(* IEC 61131-3 sources: beedance/reference (part 10) *)

// Commented out for beedance: it uses CHR_TO_STRING, which is commented out.
// FUNCTION_BLOCK TN_INPUT_EDIT_LINE
// VAR
// 	in_count : INT;
// 	in_Count_End : INT;
// 	in_CursorOffset : INT;
// 	by_Attr : BYTE;
// 	st_String : STRING;
// 	bo_Pos_Found : BOOL;
// 	st_CHAR : STRING(1);
// 	in_old_charpos : INT;
// END_VAR
// VAR
// 	FB_TN_SC_WRITE : TN_SC_WRITE;
// END_VAR
// VAR_IN_OUT
// 	Xus_TN_SCREEN : us_TN_SCREEN;
// 	Xus_TN_INPUT_CONTROL_DATA : us_TN_INPUT_CONTROL_DATA;
// END_VAR
//
// (* Cursorsteuerung rücksetzen *)
// in_CursorOffset := INT#0;
//
// IF Xus_TN_INPUT_CONTROL_DATA.bo_Focus = TRUE THEN
//
// 	(* Texteingabe erkannt ? *)
// 	IF Xus_TN_INPUT_CONTROL_DATA.by_Input_ASCII_Code > BYTE#0 THEN
//
// 		IF (Xus_TN_INPUT_CONTROL_DATA.bo_Input_Only_Num = TRUE AND Xus_TN_INPUT_CONTROL_DATA.bo_Input_ASCII_IsNum = TRUE)
// 			OR (Xus_TN_INPUT_CONTROL_DATA.bo_Input_Only_Num = FALSE) THEN
//
// 			(* ASCII Wert in einen String wandeln *)
// 			st_CHAR := CHR_TO_STRING(C:=Xus_TN_INPUT_CONTROL_DATA.by_Input_ASCII_Code);
//
// 			(* Eingabe übernehmen *)
// 			Xus_TN_INPUT_CONTROL_DATA.st_Input_Data := REPLACE(Xus_TN_INPUT_CONTROL_DATA.st_Input_Data,
// 			st_CHAR,INT#1,Xus_TN_INPUT_CONTROL_DATA.in_Cursor_Pos);
//
// 			in_CursorOffset := INT#1;
// 			Xus_TN_INPUT_CONTROL_DATA.bo_Update_Input := TRUE;
// 		END_IF;
// 	END_IF;
//
// 	CASE BYTE_TO_INT(Xus_TN_INPUT_CONTROL_DATA.by_Input_Exten_Code) OF
//
// 	67: (* Cursor rechts gedrückt *)
// 		in_CursorOffset := INT#1;
//
// 	68: (* Cursor links gedrückt *)
// 		in_CursorOffset := -1;
//
// 	08: (* Backspace gedrückt *)
// 		Xus_TN_INPUT_CONTROL_DATA.st_Input_Data := REPLACE(Xus_TN_INPUT_CONTROL_DATA.st_Input_Data, ' ', 1,Xus_TN_INPUT_CONTROL_DATA.in_Cursor_Pos);
// 		Xus_TN_INPUT_CONTROL_DATA.bo_Update_Input := TRUE;
// 		in_CursorOffset := -1;
//
// 	13: (* Enter-Taste gedrückt *)
// 		IF LEN(Xus_TN_INPUT_CONTROL_DATA.st_Input_Mask) > INT#00 THEN
// 			(* Eingabestring übernehmen *)
// 			Xus_TN_INPUT_CONTROL_DATA.st_Input_String := Xus_TN_INPUT_CONTROL_DATA.st_Input_Data;
//
// 			(* Eingabestring -> links und rechts Leerzeichen entfernen *)
// 			Xus_TN_INPUT_CONTROL_DATA.st_Input_String := TRIME(str:=Xus_TN_INPUT_CONTROL_DATA.st_Input_String);
// 			Xus_TN_INPUT_CONTROL_DATA.bo_Input_Entered := TRUE;
//
// 			(* neue Eingabe vorbereiten *)
// 			Xus_TN_INPUT_CONTROL_DATA.st_Input_Data := Xus_TN_INPUT_CONTROL_DATA.st_Input_Mask;
//
// 			Xus_TN_INPUT_CONTROL_DATA.in_Cursor_Pos := INT#1;
// 			Xus_TN_INPUT_CONTROL_DATA.bo_Update_Input := TRUE;
//
// 			(* suche erstes Position in Eingabemaske *)
// 			st_CHAR := MID(Xus_TN_INPUT_CONTROL_DATA.st_Input_Mask,1,Xus_TN_INPUT_CONTROL_DATA.in_Cursor_Pos);
// 			IF st_CHAR <> ' ' THEN
// 				(* nächsten Eingabeposition suchen *)
// 				in_CursorOffset := INT#1;
// 			END_IF;
// 		END_IF;
// 	END_CASE;
// END_IF;
//
// (* Cursor richtung rechts bewegen                                   *)
// IF (in_CursorOffset > INT#0) OR (Xus_TN_INPUT_CONTROL_DATA.in_Cursor_Pos = INT#0) THEN
// 	bo_Pos_Found := FALSE;
//
// 	in_Count := Xus_TN_INPUT_CONTROL_DATA.in_Cursor_Pos + INT#1;
// 	in_Count_End := LEN(Xus_TN_INPUT_CONTROL_DATA.st_Input_Mask);
//
// 	WHILE (in_count <= in_Count_End) AND (bo_Pos_Found = FALSE) DO
//
// 		st_CHAR := MID(Xus_TN_INPUT_CONTROL_DATA.st_Input_Mask,1,in_count);
// 		IF st_CHAR = ' ' THEN
// 			Xus_TN_INPUT_CONTROL_DATA.in_Cursor_Pos := in_count;
// 			Xus_TN_INPUT_CONTROL_DATA.bo_Update_Input := TRUE;
// 			bo_Pos_Found := TRUE;
// 		END_IF;
//
// 		in_count := in_count + INT#1;
//
// 	END_WHILE;
// END_IF;
//
// (* Cursor richtung links bewegen *)
// IF in_CursorOffset < INT#0 THEN
// 	bo_Pos_Found := FALSE;
//
// 	in_Count     := Xus_TN_INPUT_CONTROL_DATA.in_Cursor_Pos - INT#01;
// 	in_Count_End := INT#1;
//
// 	WHILE (in_count >= in_Count_End) AND (bo_Pos_Found = FALSE) DO
//
// 		st_CHAR := MID(Xus_TN_INPUT_CONTROL_DATA.st_Input_Mask,1,in_count);
// 		IF st_CHAR = ' ' THEN
// 			Xus_TN_INPUT_CONTROL_DATA.in_Cursor_Pos := in_count;
// 			Xus_TN_INPUT_CONTROL_DATA.bo_Update_Input := TRUE;
// 			bo_Pos_Found := TRUE;
// 		END_IF;
//
// 		in_count := in_count - INT#1;
// 	END_WHILE;
// END_IF;
//
// (* maximale Cursorposition ? *)
// IF Xus_TN_INPUT_CONTROL_DATA.in_Cursor_Pos > LEN(Xus_TN_INPUT_CONTROL_DATA.st_Input_Data) THEN
// 	Xus_TN_INPUT_CONTROL_DATA.in_Cursor_Pos := LEN(Xus_TN_INPUT_CONTROL_DATA.st_Input_Data);
// 	Xus_TN_INPUT_CONTROL_DATA.bo_Update_Input := TRUE;
// END_IF;
//
// (* minimale Cursorposition ? *)
// IF Xus_TN_INPUT_CONTROL_DATA.in_Cursor_Pos < INT#1 THEN
// 	Xus_TN_INPUT_CONTROL_DATA.in_Cursor_Pos := INT#1;
// 	Xus_TN_INPUT_CONTROL_DATA.bo_Update_Input := TRUE;
// END_IF;
//
// (* Aktualisierung der Anzeige *)
// IF (Xus_TN_INPUT_CONTROL_DATA.bo_Update_Input = TRUE) OR (Xus_TN_INPUT_CONTROL_DATA.bo_Update_All = TRUE) THEN
//
// 	(* Title-Text ausgeben *)
// 	IF (Xus_TN_INPUT_CONTROL_DATA.bo_Update_All = TRUE) THEN
//
// 		IF (Xus_TN_INPUT_CONTROL_DATA.in_Title_X_Offset = INT#00) AND (Xus_TN_INPUT_CONTROL_DATA.in_Title_Y_Offset = INT#00) THEN
// 			(* wenn Offset X,Y =0 dann Titlestring links vom Element positionieren *)
// 			FB_TN_SC_WRITE.Iin_Y := Xus_TN_INPUT_CONTROL_DATA.in_Y;
// 			FB_TN_SC_WRITE.Iin_X := Xus_TN_INPUT_CONTROL_DATA.in_X - LEN(Xus_TN_INPUT_CONTROL_DATA.st_Title_String);
// 		ELSE
// 			(* Title-Text durch Row, Color-Offset ausgeben *)
// 			FB_TN_SC_WRITE.Iin_Y := Xus_TN_INPUT_CONTROL_DATA.in_Y + Xus_TN_INPUT_CONTROL_DATA.in_Title_Y_Offset;
// 			FB_TN_SC_WRITE.Iin_X := Xus_TN_INPUT_CONTROL_DATA.in_X + Xus_TN_INPUT_CONTROL_DATA.in_Title_X_Offset;
// 		END_IF;
//
// 		(* Title-Text durch Row, Color-Offset ausgeben *)
// 		FB_TN_SC_WRITE(	Iby_ATTR := Xus_TN_INPUT_CONTROL_DATA.by_Title_Attr,
// 						Ist_STRING := Xus_TN_INPUT_CONTROL_DATA.st_Title_String,
// 						Xus_TN_SCREEN := Xus_TN_SCREEN);
// 	END_IF;
//
// 	(* Eingabetext ausgeben *)
// 	IF (Xus_TN_INPUT_CONTROL_DATA.bo_Input_Hidden = TRUE) THEN
//
// 		st_String := '';
//
// 		IF LEN(Xus_TN_INPUT_CONTROL_DATA.st_Input_Data) = LEN(Xus_TN_INPUT_CONTROL_DATA.st_Input_Mask) THEN
// 			(* Eingabemodus: HIDDEN *)
// 			FOR in_count := 1 TO LEN(Xus_TN_INPUT_CONTROL_DATA.st_Input_Data) DO
//
// 				(* Zeichen aus Eingabemaske lesen *)
// 				st_CHAR := MID(Xus_TN_INPUT_CONTROL_DATA.st_Input_Mask,1,in_count);
//
// 				(* Eingabe oder Maskenzeichen ausgeben *)
// 				IF st_CHAR = ' ' THEN
//
// 					(* Zeichen aus Eingabedata lesen *)
// 					st_CHAR := MID(Xus_TN_INPUT_CONTROL_DATA.st_Input_Data,1,in_count);
//
// 					IF st_CHAR = ' ' THEN
// 						(* Leerzeichen ausgeben *)
// 						st_String := CONCAT(st_String, ' ');
//
// 					ELSE
// 						(* verdecktes Zeichen ausgeben *)
// 						st_String := CONCAT(st_String, '*');
//
// 					END_IF;
//
// 				ELSE
// 					(* Zeichen aus Eingabemaske übernehmen *)
// 					st_CHAR := MID(Xus_TN_INPUT_CONTROL_DATA.st_Input_Data,1,in_count);
// 					st_String := CONCAT(st_String,st_CHAR);
//
// 				END_IF;
// 			END_FOR;
// 		END_IF;
// 	ELSE
//
// 		(* Eingabemodus: NORMAL *)
// 		st_String := Xus_TN_INPUT_CONTROL_DATA.st_Input_Data;
//
// 	END_IF;
//
// 	(* String ausgeben *)
//
// 	IF Xus_TN_INPUT_CONTROL_DATA.bo_Focus = TRUE THEN
// 		by_Attr := Xus_TN_INPUT_CONTROL_DATA.by_Attr_mF;
// 	ELSE
// 		by_Attr := Xus_TN_INPUT_CONTROL_DATA.by_Attr_oF;
// 	END_IF;
//
// 	FB_TN_SC_WRITE(	Iin_Y := Xus_TN_INPUT_CONTROL_DATA.in_Y,
// 					Iin_X := Xus_TN_INPUT_CONTROL_DATA.in_X,
// 					Iby_ATTR := by_Attr,
// 					Ist_STRING := st_String,
// 					Xus_TN_SCREEN := Xus_TN_SCREEN);
//
// 	(* Cursor auf aktuelle Position setzen *)
// 	Xus_TN_INPUT_CONTROL_DATA.in_Cursor_Y := Xus_TN_INPUT_CONTROL_DATA.in_Y;
// 	Xus_TN_INPUT_CONTROL_DATA.in_Cursor_X := Xus_TN_INPUT_CONTROL_DATA.in_X + Xus_TN_INPUT_CONTROL_DATA.in_Cursor_Pos - INT#1;
//
// 	in_old_charpos := INT#0;
//
// 	(* Update-Flag's rücksetzen *)
// 	Xus_TN_INPUT_CONTROL_DATA.bo_Update_All := FALSE;
// 	Xus_TN_INPUT_CONTROL_DATA.bo_Update_Input := FALSE;
// END_IF;
// END_FUNCTION_BLOCK

// Commented out for beedance: it uses ELEMENT_GET, which is commented out.
// FUNCTION_BLOCK TN_INPUT_MENU_BAR
// VAR
// 	FB_TN_INPUT_MENU_POPUP : TN_INPUT_MENU_POPUP;
// 	us_TN_MENU_POPUP : us_TN_MENU_POPUP;
// 	FB_TN_SC_WRITE_C : TN_SC_WRITE_C;
// END_VAR
// VAR
// 	in_ROW : INT;
// 	in_COL : INT;
// 	in_TITLE_Length : INT;
// 	st_MENU_BAR : STRING(STRING_LENGTH);
// 	st_MENU_TITLE : STRING;
// 	in_Count : INT;
// 	in_Index : INT;
// 	by_New_KeyCode : BYTE;
// 	in_Scroll_Offset : INT;
// 	by_ATTR : BYTE;
// 	bo_Reset_Position :	BOOL;
// END_VAR
// VAR_IN_OUT
// 	Xus_TN_MENU : us_TN_MENU;
// 	Xus_TN_SCREEN : us_TN_SCREEN;
// END_VAR
//
// (* sicherstellen das rechteck immer innerhalb screen positioniert wird *)
//
// IF (Xus_TN_MENU.in_State = INT#00) AND (Xus_TN_MENU.bo_Create = TRUE) THEN
// 	Xus_TN_MENU.in_State := INT#01;
// 	Xus_TN_MENU.bo_Create := FALSE;
// 	Xus_TN_MENU.in_Menu_Selected := INT#00;
// 	Xus_TN_MENU.bo_Update := TRUE;
// 	bo_Reset_Position := TRUE;
//
// 	(* Menu-Bar - Hauptmenue *)
// 	st_MENU_BAR := ELEMENT_GET(SEP:=BYTE#37,POS:=0,ELEMENT:=Xus_TN_MENU.st_MENU_TEXT);
//
// 	(* Menu-Bar - Anzahl der Elemente bestimmen *)
// 	Xus_TN_MENU.in_Menu_E_Count := ELEMENT_COUNT(SEP:=BYTE#35,ELEMENT:=st_MENU_BAR);
//
// END_IF;
//
// (* Keycode ablegen *)
// by_New_KeyCode := Xus_TN_SCREEN.by_Input_Exten_Code;
//
// (* Popup-Menu Tastensteuerung (nur Cursor oben + unten zulassen *)
// IF (by_New_KeyCode = BYTE#65) OR (by_New_KeyCode = BYTE#66) THEN
// 	us_TN_MENU_POPUP.by_Input_Exten_Code := by_New_KeyCode;
// ELSE
// 	us_TN_MENU_POPUP.by_Input_Exten_Code := BYTE#00;
// END_IF;
//
// (* Escape *)
// IF (by_New_KeyCode = BYTE#27) THEN
// 	(* Menu war inaktiv -> Escape -> Menu aktivieren *)
// 	IF (Xus_TN_MENU.in_State = INT#01) AND (Xus_TN_SCREEN.bo_Modal_Dialog = FALSE) THEN
// 		Xus_TN_MENU.in_State := INT#02;
// 		Xus_TN_MENU.bo_Update := TRUE;
// 		Xus_TN_MENU.in_Menu_Selected := INT#00;
//
// 		Xus_TN_SCREEN.bo_Menue_Bar_Dialog := TRUE;
//
// 		(* Menu war aktiv -> Escape -> Menu deaktivieren *)
// 	ELSIF (Xus_TN_MENU.in_State = INT#02) THEN
// 		us_TN_MENU_POPUP.bo_Destroy := TRUE;
// 		Xus_TN_MENU.bo_Update := TRUE;
// 		Xus_TN_MENU.in_State := INT#01;
// 		bo_Reset_Position := TRUE;
//
// 		Xus_TN_SCREEN.bo_Menue_Bar_Dialog := FALSE;
// 	END_IF;
// END_IF;
//
// (* Menu aktiv *)
// IF (Xus_TN_MENU.in_State = INT#02) THEN
//
// 	(* Return *)
// 	IF (by_New_KeyCode = BYTE#13)  THEN
// 		us_TN_MENU_POPUP.bo_Destroy := TRUE;
// 		Xus_TN_MENU.bo_Update := TRUE;
// 		Xus_TN_MENU.in_State := INT#01;
// 		bo_Reset_Position := TRUE;
// 		Xus_TN_MENU.in_Menu_Selected := (Xus_TN_MENU.in_Cur_Menu_Item * INT#10) + Xus_TN_MENU.in_Cur_Sub_Item;
// 		Xus_TN_SCREEN.by_Input_Exten_Code := BYTE#00;
//
// 		Xus_TN_SCREEN.bo_Menue_Bar_Dialog := FALSE;
//
// 		(* Destroy-Befehl -> Popup-Menu beenden *)
// 	ELSIF (Xus_TN_MENU.bo_Destroy = TRUE) THEN
// 		us_TN_MENU_POPUP.bo_Destroy := TRUE;
// 		Xus_TN_MENU.bo_Update := TRUE;
// 		Xus_TN_MENU.in_State := INT#01;
// 		bo_Reset_Position := TRUE;
// 		Xus_TN_MENU.in_Menu_Selected := INT#00;
// 		Xus_TN_SCREEN.by_Input_Exten_Code := BYTE#00;
//
// 		Xus_TN_SCREEN.bo_Menue_Bar_Dialog := FALSE;
//
// 	END_IF;
//
// 	IF (by_New_KeyCode = BYTE#67) THEN (* Cursor rechts *)
// 		in_Scroll_Offset := INT#1;
// 		Xus_TN_MENU.bo_Update := TRUE;
// 		Xus_TN_SCREEN.by_Input_Exten_Code := BYTE#00;
//
// 	ELSIF (by_New_KeyCode = BYTE#68) THEN (* Cursor links *)
// 		in_Scroll_Offset := -1;
// 		Xus_TN_MENU.bo_Update := TRUE;
// 		Xus_TN_SCREEN.by_Input_Exten_Code := BYTE#00;
// 	END_IF;
// END_IF;
//
// IF bo_Reset_Position = TRUE THEN
// 	bo_Reset_Position := FALSE;
// 	Xus_TN_MENU.in_X_SM_old := -1;
// 	Xus_TN_MENU.in_Y_SM_old := -1;
// 	Xus_TN_MENU.in_X_SM_new := -1;
// 	Xus_TN_MENU.in_Y_SM_new := -1;
// END_IF;
//
// (* POPUP-Menu updaten *)
// IF (Xus_TN_MENU.in_State > INT#00) AND (Xus_TN_MENU.bo_Update = TRUE) THEN
//
// 	Xus_TN_MENU.bo_Update := FALSE;
//
// 	in_ROW := Xus_TN_MENU.in_Y;
// 	in_COL := Xus_TN_MENU.in_X;
//
// 	(* Scrolloffset *)
// 	IF in_Scroll_Offset <> INT#00 THEN
// 		Xus_TN_MENU.in_Cur_Menu_Item := INC2(Xus_TN_MENU.in_Cur_Menu_Item,in_Scroll_Offset,1,Xus_TN_MENU.in_Menu_E_Count);
// 		in_Scroll_Offset := INT#00;
// 	ELSE
// 		(* Item = 0 und kein Scrolloffset *)
// 		IF (Xus_TN_MENU.in_Cur_Menu_Item = INT#00) THEN
// 			Xus_TN_MENU.in_Cur_Menu_Item := INT#01;
// 		END_IF;
// 	END_IF;
//
// 	(* alle Menutext zeichnen *)
// 	FOR in_Count := INT#01 TO Xus_TN_MENU.in_Menu_E_Count DO;
//
// 		(* Zeichenfarbe bestimmen *)
// 		IF (in_Count = Xus_TN_MENU.in_Cur_Menu_Item) AND (Xus_TN_MENU.in_State > INT#01 ) THEN
// 			by_ATTR := Xus_TN_MENU.by_Attr_mF;
//
// 			Xus_TN_MENU.in_Y_SM_new := in_ROW + INT#01;
// 			Xus_TN_MENU.in_X_SM_new := in_COL;
//
// 		ELSE
// 			by_ATTR := Xus_TN_MENU.by_Attr_oF;
// 		END_IF;
//
// 		st_MENU_TITLE := ELEMENT_GET(SEP:=BYTE#35,POS:=in_Count - 1,ELEMENT:=st_MENU_BAR);
//
// 		in_TITLE_Length := LEN(st_MENU_TITLE) + INT#02;
//
// 		FB_TN_SC_WRITE_C(	Iin_Y := in_ROW,
// 							Iin_X := in_COL,
// 							Iby_ATTR := by_ATTR,
// 							Iin_LENGTH := in_TITLE_Length,
// 							Iin_OPTION := INT#02,
// 							Ist_STRING := st_MENU_TITLE,
// 							Xus_TN_SCREEN := Xus_TN_SCREEN);
//
// 		in_COL := in_COL + in_TITLE_Length;
//
// 	END_FOR;
// END_IF;
//
// IF Xus_TN_MENU.in_X_SM_new <> Xus_TN_MENU.in_X_SM_old THEN
//
// 	(* SubMenu ist aktiv -> beenden                                     *)
// 	IF us_TN_MENU_POPUP.bo_Activ = TRUE THEN
// 		us_TN_MENU_POPUP.bo_Destroy := TRUE;
//
// 		(* Sub-Menu bearbeiten *)
// 		FB_TN_INPUT_MENU_POPUP(	Xus_TN_MENU_POPUP := us_TN_MENU_POPUP,
// 								Xus_TN_SCREEN := Xus_TN_SCREEN);
// 	END_IF;
//
// 	IF us_TN_MENU_POPUP.bo_Activ = FALSE THEN
// 		(* Popup-Menu zu aktuellen Menu parametrieren und ausführen         *)
// 		in_Index := Xus_TN_MENU.in_Cur_Menu_Item;
//
// 		us_TN_MENU_POPUP.in_Y := Xus_TN_MENU.in_Y_SM_new;
// 		us_TN_MENU_POPUP.in_X := Xus_TN_MENU.in_X_SM_new;
// 		us_TN_MENU_POPUP.by_Attr_mF := Xus_TN_MENU.by_Attr_mF;
// 		us_TN_MENU_POPUP.by_Attr_oF := Xus_TN_MENU.by_Attr_oF;
// 		us_TN_MENU_POPUP.st_Menu_Text := ELEMENT_GET(SEP:=BYTE#37,POS:=in_Index,ELEMENT:=Xus_TN_MENU.st_MENU_TEXT);
// 		us_TN_MENU_POPUP.bo_Create := TRUE;
//
// 		Xus_TN_MENU.in_X_SM_old := Xus_TN_MENU.in_X_SM_new;
// 		Xus_TN_MENU.in_Y_SM_old := Xus_TN_MENU.in_Y_SM_new;
//
// 	END_IF;
// END_IF;
//
// (* Popup-Menu zyklisch aufrufen *)
// FB_TN_INPUT_MENU_POPUP(	Xus_TN_MENU_POPUP := us_TN_MENU_POPUP,
// 						Xus_TN_SCREEN := Xus_TN_SCREEN);
//
// (* aktuelles Item vom Popup-Menu kopieren *)
// Xus_TN_MENU.in_Cur_Sub_Item := us_TN_MENU_POPUP.in_Cur_Item;
//
// (* Destroy-Befehl *)
// IF (Xus_TN_MENU.in_State = INT#01) THEN
// 	IF (Xus_TN_MENU.bo_Destroy = TRUE) THEN
// 		Xus_TN_MENU.in_State := INT#00;
// 		Xus_TN_MENU.bo_Destroy := FALSE;
// 		Xus_TN_MENU.in_Cur_Menu_Item := INT#00;
// 		Xus_TN_MENU.in_Cur_Sub_Item := INT#00;
// 	END_IF;
// END_IF;
// END_FUNCTION_BLOCK

// Commented out for beedance: it uses ELEMENT_COUNT, which is commented out.
// FUNCTION_BLOCK TN_INPUT_MENU_POPUP
// VAR
// 	FB_TN_SC_AREA_SAVE : TN_SC_AREA_SAVE;
// 	FB_TN_SC_AREA_RESTORE : TN_SC_AREA_RESTORE;
// 	FB_TN_SC_LINE : TN_SC_LINE;
// 	FB_TN_SC_ADD_SHADOW : TN_SC_ADD_SHADOW;
// 	FB_TN_SC_BOX : TN_SC_BOX;
// 	FB_TN_SC_WRITE_C : TN_SC_WRITE_C;
// END_VAR
// VAR
// 	in_ROW : INT;
// 	in_ROWS : INT;
// 	in_COL : INT;
// 	in_COLS : INT;
// 	in_index : INT;
// 	in_Count : INT;
// 	in_Scroll_Offset : INT;
// 	by_ATTR : BYTE;
// END_VAR
// VAR_IN_OUT
// 	Xus_TN_MENU_POPUP : us_TN_MENU_POPUP;
// 	Xus_TN_SCREEN : us_TN_SCREEN;
// END_VAR
//
// (* sicherstellen das rechteck immer innerhalb screen positioniert wird *)
//
// IF (Xus_TN_MENU_POPUP.bo_Activ = FALSE) AND (Xus_TN_MENU_POPUP.bo_Create = TRUE) THEN
// 	Xus_TN_MENU_POPUP.bo_Activ := TRUE;
// 	Xus_TN_MENU_POPUP.bo_Create := FALSE;
// 	Xus_TN_MENU_POPUP.bo_Destroy := FALSE;
// 	Xus_TN_MENU_POPUP.bo_Update := TRUE;
//
//   (* Sub-Menu-Texte *)
//
// 	Xus_TN_MENU_POPUP.in_Menu_E_Count := ELEMENT_COUNT(SEP:=BYTE#35,ELEMENT:=Xus_TN_MENU_POPUP.st_Menu_Text);
//
// 	(* Anzahl Zeilen (Sub-Menu-Texte) bestimmen *)
// 	Xus_TN_MENU_POPUP.in_Rows := Xus_TN_MENU_POPUP.in_Menu_E_Count;
//
// 	(* längsten Sub-Menu-Text suchen *)
// 	Xus_TN_MENU_POPUP.in_Cols := INT#00;
//
// 	FOR in_Count := INT#01 TO Xus_TN_MENU_POPUP.in_Rows DO;
// 		Xus_TN_MENU_POPUP.in_Cols:=MAX(LEN(ELEMENT_GET(SEP:=BYTE#35,POS:=in_Count - 1,ELEMENT:=Xus_TN_MENU_POPUP.st_Menu_Text)),Xus_TN_MENU_POPUP.in_Cols);
// 	END_FOR;
//
// 	(* Horizontale Position überprüfen und korrigieren *)
// 	IF (Xus_TN_MENU_POPUP.in_X + Xus_TN_MENU_POPUP.in_Cols) > INT#75 THEN
// 		Xus_TN_MENU_POPUP.in_X := INT#79 - Xus_TN_MENU_POPUP.in_Cols - INT#04;
// 	END_IF;
//
//   (* Vertikale Position überprüfen und korrigieren *)
// 	IF (Xus_TN_MENU_POPUP.in_Y + Xus_TN_MENU_POPUP.in_ROWS) > INT#21 THEN
// 		Xus_TN_MENU_POPUP.in_Y := INT#23 - Xus_TN_MENU_POPUP.in_ROWS - INT#2;
// 	END_IF;
//
// 	Xus_TN_SCREEN.bo_Modal_Dialog := TRUE;
//
// 	(* Hintergrund sichern *)
// 	FB_TN_SC_AREA_SAVE(	Iin_X1 := Xus_TN_MENU_POPUP.in_X,
// 									Iin_Y1 := Xus_TN_MENU_POPUP.in_Y,
// 									Iin_X2 := Xus_TN_MENU_POPUP.in_X + Xus_TN_MENU_POPUP.in_Cols + INT#04,
// 									Iin_Y2 := Xus_TN_MENU_POPUP.in_Y + Xus_TN_MENU_POPUP.in_Rows + INT#02,
// 									Xus_TN_SCREEN := Xus_TN_SCREEN);
//
// 	(* Rahmen für Submenu zeichnen *)
// 	FB_TN_SC_BOX(	Iin_X1 := Xus_TN_MENU_POPUP.in_X,
// 					Iin_Y1 := Xus_TN_MENU_POPUP.in_Y,
// 					Iin_X2 := Xus_TN_MENU_POPUP.in_X + Xus_TN_MENU_POPUP.in_Cols + INT#03,
// 					Iin_Y2 := Xus_TN_MENU_POPUP.in_Y + Xus_TN_MENU_POPUP.in_Rows + INT#01,
// 					Iby_FILL := BYTE#32, (* Füllung *)
// 					Iin_BORDER := INT#01, (* Single-Line Border *)
// 					Iby_ATTR := Xus_TN_MENU_POPUP.by_Attr_oF,
// 					Xus_TN_SCREEN := Xus_TN_SCREEN);
//
// 	(* Shadow für Submenu zeichnen *)
// 	FB_TN_SC_ADD_SHADOW(Iin_X1 := Xus_TN_MENU_POPUP.in_X + INT#1,
// 						Iin_Y1 := Xus_TN_MENU_POPUP.in_Y + INT#1,
// 						Iin_X2 := Xus_TN_MENU_POPUP.in_X + Xus_TN_MENU_POPUP.in_Cols + INT#04,
// 						Iin_Y2 := Xus_TN_MENU_POPUP.in_Y + Xus_TN_MENU_POPUP.in_Rows + INT#02,
// 						Iin_OPTION := INT#00,
// 						Xus_TN_SCREEN := Xus_TN_SCREEN);
//
// 	(* Parameter laden *)
// 	in_COL := Xus_TN_MENU_POPUP.in_X;
// 	in_ROW := Xus_TN_MENU_POPUP.in_Y;
// 	in_ROWS := Xus_TN_MENU_POPUP.in_Rows;
// 	in_COLS := Xus_TN_MENU_POPUP.in_Cols;
//
// 	(* Trennlinien zeichnen *)
// 	in_COLS := in_COLS + INT#02; (* Text um 2 Zeichen verlängern *)
//
// 	FOR in_Count := INT#01 TO Xus_TN_MENU_POPUP.in_Menu_E_Count DO;
// 		in_ROW := in_ROW + INT#01;
//
// 		IF ELEMENT_GET(SEP:=BYTE#35,POS:=in_Count - 1,ELEMENT:=Xus_TN_MENU_POPUP.st_Menu_Text) = '-' THEN
//
// 			FB_TN_SC_LINE(	Iin_Y1 := in_ROW,
// 							Iin_X1 := in_COL,
// 							Iin_Y2 := in_ROW,
// 							Iin_X2 := in_COL + in_COLS + INT#01,
// 							Iby_ATTR := Xus_TN_MENU_POPUP.by_Attr_oF,
// 							Iby_BORDER := BYTE#01,
// 							Xus_TN_SCREEN := Xus_TN_SCREEN);
// 		END_IF;
// 	END_FOR;
// END_IF;
//
// IF (Xus_TN_MENU_POPUP.bo_Activ = TRUE) THEN
//
// 	CASE BYTE_TO_INT(Xus_TN_MENU_POPUP.by_Input_Exten_Code) OF
//
// 	65: (* Cursor oben *)
// 		in_Scroll_Offset := -1;
// 		Xus_TN_MENU_POPUP.bo_Update := TRUE;
//
// 	66: (* Cursor unten *)
// 		in_Scroll_Offset := 1;
// 		Xus_TN_MENU_POPUP.bo_Update := TRUE;
//
// 	13:  (* Enter *)
// 		Xus_TN_MENU_POPUP.bo_Destroy := TRUE;
//
// 	27:  (* Escape*)
// 		Xus_TN_MENU_POPUP.bo_Destroy := TRUE;
// 		Xus_TN_MENU_POPUP.in_Cur_Item := INT#00;
//
// 	67..68: (* Cursor links oder rechts *)
// 		Xus_TN_MENU_POPUP.bo_Destroy := TRUE;
// 		Xus_TN_MENU_POPUP.in_Cur_Item := INT#00;
//
// 	END_CASE;
// END_IF;
//
// (* POPUP-Menu updaten *)
// IF (Xus_TN_MENU_POPUP.bo_Activ = TRUE) AND (Xus_TN_MENU_POPUP.bo_Update = TRUE) THEN
//
// 	Xus_TN_MENU_POPUP.bo_Update := FALSE;
//
// 	(* überprüfung + nächstes anwählbares Sub-Menu suchen *)
// 	in_index := Xus_TN_MENU_POPUP.in_Cur_Item;
//
// 	IF (in_index < INT#01) OR (in_index > Xus_TN_MENU_POPUP.in_Menu_E_Count) THEN
// 		in_Scroll_Offset := INT#01;
// 		in_index := Xus_TN_MENU_POPUP.in_Menu_E_Count;
// 	END_IF;
//
// 	(* aktueller Index steht auf Trennzeichen -> ändern *)
// 	IF ELEMENT_GET(SEP:=BYTE#35,POS:=in_index-1,ELEMENT:=Xus_TN_MENU_POPUP.st_Menu_Text) = '-' THEN
// 		in_Scroll_Offset := INT#01;
// 	END_IF;
//
// 	(* Scroll-Offset *)
// 	IF in_Scroll_Offset <> INT#00 THEN
//
// 		FOR in_Count := INT#01 TO Xus_TN_MENU_POPUP.in_Menu_E_Count DO;
//
// 			in_index:=INC2(in_index,in_Scroll_Offset,1,Xus_TN_MENU_POPUP.in_Menu_E_Count);
//
// 			IF ELEMENT_GET(SEP:=BYTE#35,POS:=in_index - 1,ELEMENT:=Xus_TN_MENU_POPUP.st_Menu_Text) <> '-' THEN
// 				EXIT;
// 			END_IF;
//
// 		END_FOR;
// 	END_IF;
//
// 	Xus_TN_MENU_POPUP.in_Cur_Item := in_index;
// 	in_Scroll_Offset := INT#00;
//
// 	(* Parameter laden *)
// 	in_COL  := Xus_TN_MENU_POPUP.in_X;
// 	in_ROW  := Xus_TN_MENU_POPUP.in_Y;
// 	in_ROWS := Xus_TN_MENU_POPUP.in_Rows;
// 	in_COLS := Xus_TN_MENU_POPUP.in_Cols;
//
// 	(* SUB-MENU-Titel ausgeben *)
// 	in_COLS := in_COLS + INT#02; (* Text um 2 Zeichen verlängern *)
//
// 	FOR in_Count := INT#01 TO Xus_TN_MENU_POPUP.in_Menu_E_Count DO;
//
// 		in_ROW := in_ROW + INT#01;
//
// 		(* Zeichenfarbe bestimmen *)
// 		IF in_Count = Xus_TN_MENU_POPUP.in_Cur_Item THEN
// 			by_ATTR := Xus_TN_MENU_POPUP.by_Attr_mF;
// 		ELSE
// 			by_ATTR := Xus_TN_MENU_POPUP.by_Attr_oF;
// 		END_IF;
//
// 		FB_TN_SC_WRITE_C.Ist_STRING := ELEMENT_GET(SEP:=BYTE#35,POS:=in_Count - 1,ELEMENT:=Xus_TN_MENU_POPUP.st_Menu_Text);
//
// 		IF FB_TN_SC_WRITE_C.Ist_STRING <> '-' THEN
//
// 			FB_TN_SC_WRITE_C(	Iin_Y := in_ROW,
// 								Iin_X := in_COL + INT#01,
// 								Iby_ATTR := by_ATTR,
// 								Iin_LENGTH := in_COLS,
// 								Iin_OPTION := INT#02, (* Center *)
// 								Xus_TN_SCREEN := Xus_TN_SCREEN);
// 		END_IF;
// 	END_FOR;
// END_IF;
//
// (* POPUP-Menu entfernen (Destroy) *)
// IF (Xus_TN_MENU_POPUP.bo_Activ = TRUE) AND (Xus_TN_MENU_POPUP.bo_Destroy = TRUE) THEN
//
// 	Xus_TN_MENU_POPUP.bo_Destroy := FALSE;
// 	Xus_TN_MENU_POPUP.bo_Activ := FALSE;
//
// 	(* alten Hintergrund aus Speicher wiederherstellen *)
// 	FB_TN_SC_AREA_RESTORE(Xus_TN_SCREEN := Xus_TN_SCREEN);
//
// 	Xus_TN_SCREEN.bo_Modal_Dialog := FALSE;
// END_IF;
// END_FUNCTION_BLOCK

// Commented out for beedance: it uses TN_INPUT_MENU_POPUP, which is commented out.
// FUNCTION_BLOCK TN_INPUT_SELECT_POPUP
// VAR
// 	in_index : INT;
// 	in_Element_Count : INT;
// 	by_Cur_Key : BYTE;
// 	by_Attr : BYTE;
// 	st_String : STRING;
// END_VAR
// VAR
// 	us_TN_MENU_POPUP : us_TN_MENU_POPUP;
// 	FB_TN_INPUT_MENU_POPUP : TN_INPUT_MENU_POPUP;
// 	FB_TN_SC_WRITE : TN_SC_WRITE;
// END_VAR
// VAR_IN_OUT
// 	Xus_TN_SCREEN : us_TN_SCREEN;
// 	Xus_TN_INPUT_CONTROL_DATA : us_TN_INPUT_CONTROL_DATA;
// END_VAR
//
// (* Benutzereingabe auswerten -> Selektion Text n *)
// IF (Xus_TN_INPUT_CONTROL_DATA.bo_Focus = TRUE) THEN
//
// 	by_Cur_Key := Xus_TN_INPUT_CONTROL_DATA.by_Input_Exten_Code;
//
// 	IF (us_TN_MENU_POPUP.bo_Activ = FALSE) THEN
// 		us_TN_MENU_POPUP.by_Input_Exten_Code := BYTE#00;
//
// 		(* Return-Taste auswerten *)
// 		IF (by_Cur_Key = BYTE#13) THEN
// 			(* Popup-Menu parameter übergeben *)
// 			us_TN_MENU_POPUP.in_Y := Xus_TN_INPUT_CONTROL_DATA.in_Y;
// 			us_TN_MENU_POPUP.in_X := Xus_TN_INPUT_CONTROL_DATA.in_X;
// 			us_TN_MENU_POPUP.by_Attr_mF := Xus_TN_INPUT_CONTROL_DATA.by_Attr_mF;
// 			us_TN_MENU_POPUP.by_Attr_oF := Xus_TN_INPUT_CONTROL_DATA.by_Attr_oF;
// 			us_TN_MENU_POPUP.st_Menu_Text := Xus_TN_INPUT_CONTROL_DATA.st_Input_Data;
// 			us_TN_MENU_POPUP.bo_Create := TRUE;
// 			us_TN_MENU_POPUP.in_Cur_Item := INT#00;
// 		END_IF;
//
// 		IF (us_TN_MENU_POPUP.in_Cur_Item > INT#00) THEN
// 			Xus_TN_INPUT_CONTROL_DATA.in_selected := us_TN_MENU_POPUP.in_Cur_Item;
// 			Xus_TN_INPUT_CONTROL_DATA.bo_Input_Entered := TRUE;
// 			Xus_TN_INPUT_CONTROL_DATA.bo_Update_Input := TRUE;
// 			us_TN_MENU_POPUP.in_Cur_Item := INT#00;
// 		END_IF;
//
// 	ELSE
// 		us_TN_MENU_POPUP.by_Input_Exten_Code := by_Cur_Key;
// 	END_IF;
//
// 	(* Popup-Menu zyklisch aufrufen *)
// 	FB_TN_INPUT_MENU_POPUP(Xus_TN_MENU_POPUP := us_TN_MENU_POPUP, Xus_TN_SCREEN := Xus_TN_SCREEN);
//
// END_IF;
//
// (* Aktualisierung der Anzeige *)
// IF (Xus_TN_INPUT_CONTROL_DATA.bo_Update_Input = TRUE) OR (Xus_TN_INPUT_CONTROL_DATA.bo_Update_All = TRUE) THEN
//
// 	(* Title-Text ausgeben *)
// 	IF Xus_TN_INPUT_CONTROL_DATA.bo_Update_All = TRUE THEN
//
// 		IF (Xus_TN_INPUT_CONTROL_DATA.in_Title_X_Offset = INT#00) AND (Xus_TN_INPUT_CONTROL_DATA.in_Title_Y_Offset = INT#00) THEN
// 			(* wenn Offset X,Y =0 dann Titlestring links vom Element positionieren *)
// 			FB_TN_SC_WRITE.Iin_Y := Xus_TN_INPUT_CONTROL_DATA.in_Y;
// 			FB_TN_SC_WRITE.Iin_X := Xus_TN_INPUT_CONTROL_DATA.in_X - LEN(Xus_TN_INPUT_CONTROL_DATA.st_Title_String);
//
// 		ELSE
// 			(* Title-Text durch Row, Color-Offset ausgeben *)
// 			FB_TN_SC_WRITE.Iin_Y := Xus_TN_INPUT_CONTROL_DATA.in_Y + Xus_TN_INPUT_CONTROL_DATA.in_Title_Y_Offset;
// 			FB_TN_SC_WRITE.Iin_X := Xus_TN_INPUT_CONTROL_DATA.in_X + Xus_TN_INPUT_CONTROL_DATA.in_Title_X_Offset;
// 		END_IF;
//
// 		(* Title-Text durch Row, Color-Offset ausgeben *)
// 		FB_TN_SC_WRITE(	Iby_ATTR := Xus_TN_INPUT_CONTROL_DATA.by_Title_Attr,
// 						Ist_STRING := Xus_TN_INPUT_CONTROL_DATA.st_Title_String,
// 						Xus_TN_SCREEN := Xus_TN_SCREEN);
// 	END_IF;
//
// 	in_Element_Count := ELEMENT_COUNT(SEP:=BYTE#35,ELEMENT:=Xus_TN_INPUT_CONTROL_DATA.st_Input_Data);
//
// 	IF in_Element_Count > INT#00 THEN
//
// 		Xus_TN_INPUT_CONTROL_DATA.in_selected:=LIMIT(1,Xus_TN_INPUT_CONTROL_DATA.in_selected,in_Element_Count);
//
// 		in_index := Xus_TN_INPUT_CONTROL_DATA.in_selected;
//
// 		st_String := ELEMENT_GET(SEP:=BYTE#35,POS:=in_index - 1,ELEMENT:=Xus_TN_INPUT_CONTROL_DATA.st_Input_Data);
//
// 		st_String:= FIX(str:=st_String,
// 						L:=LEN(Xus_TN_INPUT_CONTROL_DATA.st_Input_Mask),
// 						C:=BYTE#32,
// 						M:=Xus_TN_INPUT_CONTROL_DATA.in_Input_Option);
//
// 		Xus_TN_INPUT_CONTROL_DATA.st_Input_String := st_String;
//
// 		IF Xus_TN_INPUT_CONTROL_DATA.bo_Focus = TRUE THEN
// 			by_Attr := Xus_TN_INPUT_CONTROL_DATA.by_Attr_mF;
// 		ELSE
// 			by_Attr := Xus_TN_INPUT_CONTROL_DATA.by_Attr_oF;
// 		END_IF;
//
// 		FB_TN_SC_WRITE(	Iin_X := Xus_TN_INPUT_CONTROL_DATA.in_X,
// 								Iin_Y := Xus_TN_INPUT_CONTROL_DATA.in_Y,
// 								Iby_ATTR := by_Attr,
// 								Ist_STRING := st_String,
// 								Xus_TN_SCREEN := Xus_TN_SCREEN );
// 	END_IF;
//
// 	(* Cursor auf aktuelle Position setzen *)
// 	Xus_TN_INPUT_CONTROL_DATA.in_Cursor_X := Xus_TN_INPUT_CONTROL_DATA.in_X;
// 	Xus_TN_INPUT_CONTROL_DATA.in_Cursor_Y := Xus_TN_INPUT_CONTROL_DATA.in_Y;
//
// 	(* Update-Flag's rücksetzen *)
// 	Xus_TN_INPUT_CONTROL_DATA.bo_Update_All   := FALSE;
// 	Xus_TN_INPUT_CONTROL_DATA.bo_Update_Input := FALSE;
//
// END_IF;
// END_FUNCTION_BLOCK

// Commented out for beedance: it uses ELEMENT_COUNT, which is commented out.
// FUNCTION_BLOCK TN_INPUT_SELECT_TEXT
// VAR
// 	in_count : INT;
// 	by_Attr : BYTE;
// 	st_String : STRING;
// END_VAR
// VAR
// 	FB_TN_SC_WRITE : TN_SC_WRITE;
// END_VAR
// VAR_IN_OUT
// 	Xus_TN_SCREEN : us_TN_SCREEN;
// 	Xus_TN_INPUT_CONTROL_DATA : us_TN_INPUT_CONTROL_DATA;
// END_VAR
//
// (* Benutzereingabe auswerten -> Selektion Text n *)
// IF Xus_TN_INPUT_CONTROL_DATA.bo_Focus = TRUE THEN
//
// (* Leertaste-Taste auswerten *)
// 	IF Xus_TN_INPUT_CONTROL_DATA.by_Input_ASCII_Code = BYTE#32 THEN
// 		Xus_TN_INPUT_CONTROL_DATA.in_selected := Xus_TN_INPUT_CONTROL_DATA.in_selected + INT#01;
// 		Xus_TN_INPUT_CONTROL_DATA.bo_Update_Input := TRUE;
// 	END_IF;
//
// 	(* Return-Taste auswerten *)
// 	IF Xus_TN_INPUT_CONTROL_DATA.by_Input_Exten_Code = BYTE#13 THEN
// 		Xus_TN_INPUT_CONTROL_DATA.bo_Input_Entered := TRUE;
// 	END_IF;
//
// END_IF;
//
// (* Aktualisierung der Anzeige *)
// IF (Xus_TN_INPUT_CONTROL_DATA.bo_Update_Input = TRUE) OR (Xus_TN_INPUT_CONTROL_DATA.bo_Update_All = TRUE) THEN
//
// 	(* Title-Text ausgeben *)
// 	IF Xus_TN_INPUT_CONTROL_DATA.bo_Update_All = TRUE THEN
//
// 		IF (Xus_TN_INPUT_CONTROL_DATA.in_Title_X_Offset = INT#00) AND (Xus_TN_INPUT_CONTROL_DATA.in_Title_Y_Offset = INT#00) THEN
// 			(* wenn Offset X,Y =0 dann Titlestring links vom Element positionieren *)
// 			FB_TN_SC_WRITE.Iin_Y := Xus_TN_INPUT_CONTROL_DATA.in_Y;
// 			FB_TN_SC_WRITE.Iin_X := Xus_TN_INPUT_CONTROL_DATA.in_X - LEN(Xus_TN_INPUT_CONTROL_DATA.st_Title_String);
//
// 		ELSE
// 			(* Title-Text durch Row, Color-Offset ausgeben *)
// 			FB_TN_SC_WRITE.Iin_Y := Xus_TN_INPUT_CONTROL_DATA.in_Y + Xus_TN_INPUT_CONTROL_DATA.in_Title_Y_Offset;
// 			FB_TN_SC_WRITE.Iin_X := Xus_TN_INPUT_CONTROL_DATA.in_X + Xus_TN_INPUT_CONTROL_DATA.in_Title_X_Offset;
// 		END_IF;
//
// 		(* Title-Text durch Row, Color-Offset ausgeben *)
// 		FB_TN_SC_WRITE(	Iby_ATTR := Xus_TN_INPUT_CONTROL_DATA.by_Title_Attr,
// 						Ist_STRING := Xus_TN_INPUT_CONTROL_DATA.st_Title_String,
// 						Xus_TN_SCREEN := Xus_TN_SCREEN);
//
// 	END_IF;
//
// 	(* Eingabezeile verarbeiten *)
//
// 	(* Anzahl der Elemente bestimmen *)
// 	in_count := ELEMENT_COUNT(SEP:=BYTE#35,ELEMENT:=Xus_TN_INPUT_CONTROL_DATA.st_Input_Data);
//
// 	IF in_Count > INT#00 THEN
//
// 		IF Xus_TN_INPUT_CONTROL_DATA.in_selected < INT#1 THEN
// 			Xus_TN_INPUT_CONTROL_DATA.in_selected := INT#01;
// 		END_IF;
//
// 		IF Xus_TN_INPUT_CONTROL_DATA.in_selected > in_count THEN
// 			Xus_TN_INPUT_CONTROL_DATA.in_selected := INT#01;
// 		END_IF;
//
// 		st_String := ELEMENT_GET(SEP:=BYTE#35,POS:=Xus_TN_INPUT_CONTROL_DATA.in_selected - 1,ELEMENT:=Xus_TN_INPUT_CONTROL_DATA.st_Input_Data);
//
// 		st_String := FIX(	str:=st_String,
// 							L:=LEN(Xus_TN_INPUT_CONTROL_DATA.st_Input_Mask),
// 							C:=BYTE#32,
// 							M:=Xus_TN_INPUT_CONTROL_DATA.in_Input_Option);
//
// 		Xus_TN_INPUT_CONTROL_DATA.st_Input_String := st_String;
//
// 		IF Xus_TN_INPUT_CONTROL_DATA.bo_Focus = TRUE THEN
// 			by_Attr := Xus_TN_INPUT_CONTROL_DATA.by_Attr_mF;
// 		ELSE
// 			by_Attr := Xus_TN_INPUT_CONTROL_DATA.by_Attr_oF;
// 		END_IF;
//
// 		FB_TN_SC_WRITE(	Iin_Y := Xus_TN_INPUT_CONTROL_DATA.in_Y,
// 						Iin_X := Xus_TN_INPUT_CONTROL_DATA.in_X,
// 						Iby_ATTR := by_Attr,
// 						Ist_STRING := st_String,
// 						Xus_TN_SCREEN := Xus_TN_SCREEN);
// 	END_IF;
//
// 	(* Cursor auf aktuelle Position setzen *)
// 	Xus_TN_INPUT_CONTROL_DATA.in_Cursor_Y := Xus_TN_INPUT_CONTROL_DATA.in_Y;
// 	Xus_TN_INPUT_CONTROL_DATA.in_Cursor_X := Xus_TN_INPUT_CONTROL_DATA.in_X;
//
// 	(* Update-Flag's rücksetzen *)
// 	Xus_TN_INPUT_CONTROL_DATA.bo_Update_All := FALSE;
// 	Xus_TN_INPUT_CONTROL_DATA.bo_Update_Input := FALSE;
//
// END_IF;
// END_FUNCTION_BLOCK

FUNCTION_BLOCK TN_RECEIVE
VAR_IN_OUT
	R_BUF :	NETWORK_BUFFER;
	Xus_TN_SCREEN : us_TN_SCREEN;
END_VAR
VAR
	REQ_Size : UINT;
	REQ1 : BYTE;
	REQ2 : BYTE;
	REQ3 : BYTE;
END_VAR

(* Datenempfang auswertung *)
Xus_TN_SCREEN.by_Input_ASCII_Code := BYTE#00;
Xus_TN_SCREEN.by_Input_Exten_Code := BYTE#00;

IF R_BUF.SIZE > UINT#0 THEN
	(* empfangene Daten auswerten *)
	REQ_Size := R_BUF.SIZE;
	REQ1 := R_BUF.BUFFER[0];
	REQ2 := R_BUF.BUFFER[1];
	REQ3 := R_BUF.BUFFER[2];

	IF REQ1 = BYTE#27 AND REQ_Size >= UINT#3 THEN (* Escape *)
		IF REQ2 = BYTE#91 THEN (* Cursor code *)
			IF (REQ3 >= BYTE#65 AND REQ3 <= BYTE#68) OR (REQ3 = BYTE#72) OR (REQ3 = BYTE#75) THEN (* 65..68 = Cursor o,u,r,l / 72 = POS1 / 75 = ENDE *)
				Xus_TN_SCREEN.by_Input_Exten_Code := REQ3;
			END_IF;
		ELSIF REQ2 = BYTE#79 THEN (* Sondertasten F1/F2/F3/F4 *)
			IF REQ3 >= BYTE#80 AND REQ3 <= BYTE#83 THEN
				Xus_TN_SCREEN.by_Input_Exten_Code := REQ3;
			END_IF;
		END_IF;
	ELSIF REQ1 >= BYTE#32 AND REQ1 <= BYTE#126 THEN
		Xus_TN_SCREEN.by_Input_ASCII_Code := REQ1;
		Xus_TN_SCREEN.bo_Input_ASCII_IsNum := ISC_NUM(REQ1); (* Auswertung auf Zahleneingabe *)
	ELSIF REQ1 = BYTE#8 OR REQ1 = BYTE#9 OR REQ1 = BYTE#13 OR REQ1 = BYTE#27 THEN (* prüfe auf Steuerzeichen 8=Backspace / 9=Tabulator / 13=Return / 27=Escape *)
		Xus_TN_SCREEN.by_Input_Exten_Code := REQ1;
	END_IF;

	(* Empfangsbuffer Datenlänge null eintragen (Telegramm zerstören *)
	R_BUF.SIZE := UINT#00;
END_IF;
END_FUNCTION_BLOCK

FUNCTION_BLOCK TN_SC_ADD_SHADOW
VAR
	in_Offset : INT;
	in_X : INT;
	in_Y : INT;
END_VAR
VAR_INPUT
	Iin_Y1 : INT;
	Iin_X1 : INT;
	Iin_Y2 : INT;
	Iin_X2 : INT;
	Iin_OPTION : INT;
END_VAR
VAR_IN_OUT
	Xus_TN_SCREEN : us_TN_SCREEN;
END_VAR

IF TN_SC_XY2_ERROR(Iin_X1,Iin_Y1,Iin_X2,Iin_Y2) THEN RETURN; END_IF;

IF Iin_Y1 < 0 OR Iin_X1 < 0 OR Iin_Y2 < 0 OR Iin_X2 < 0 THEN RETURN; END_IF; (* min werte prüfen *)
IF Iin_Y1 > 23 OR Iin_X1 > 79 OR Iin_Y2 > 23 OR Iin_X2 > 79 THEN RETURN; END_IF; (* max werte prüfen *)

in_Offset := (Iin_Y1 * 80) + Iin_X2;

IF Iin_OPTION = INT#00 THEN
	(* Schatten durch Farbanpassung erzeugen *)
	FOR in_Y := Iin_Y1 TO Iin_Y2 DO
		Xus_TN_SCREEN.bya_COLOR[in_Offset] := TN_SC_SHADOW_ATTR(Xus_TN_SCREEN.bya_COLOR[in_Offset]);
		in_Offset := in_Offset + 80;
		Xus_TN_SCREEN.bya_Line_Update[in_Y] := TRUE; (* Zeile für Update eintragen *)
	END_FOR;
ELSE
	(* Schatten durch Farbe Schwarz und Leerzeichen erzeugen *)
	FOR in_Y := Iin_Y1 TO Iin_Y2 DO
		Xus_TN_SCREEN.bya_COLOR[in_Offset] := BYTE#00;
		Xus_TN_SCREEN.bya_CHAR[in_Offset] := BYTE#32;
		in_Offset := in_Offset + 80;
		Xus_TN_SCREEN.bya_Line_Update[in_Y] := TRUE; (* Zeile für Update eintragen *)
	END_FOR;
END_IF;

in_Offset := (Iin_Y2 * 80) + Iin_X1;

IF Iin_OPTION = INT#00 THEN
	(* Schatten durch Farbanpassung erzeugen *)
	FOR in_X  := Iin_X1 TO Iin_X2 DO
		Xus_TN_SCREEN.bya_COLOR[in_Offset] := TN_SC_SHADOW_ATTR(Xus_TN_SCREEN.bya_COLOR[in_Offset]);
		in_Offset := in_Offset + 1;
	END_FOR;
ELSE
	(* Schatten durch Farbe Schwarz und Leerzeichen erzeugen *)
	FOR in_X  := Iin_X1 TO Iin_X2 DO
		Xus_TN_SCREEN.bya_COLOR[in_Offset] := BYTE#00;
		Xus_TN_SCREEN.bya_CHAR[in_Offset] := BYTE#32;
		in_Offset := in_Offset + 1;
	END_FOR;
END_IF;
END_FUNCTION_BLOCK

FUNCTION_BLOCK TN_SC_AREA_RESTORE
VAR
	in_Offset_1 : INT;
	in_Offset_2 : INT;
	in_Y : INT;
	in_X : INT;
	in_Y1 : INT;
	in_X1 : INT;
	in_Y2 : INT;
	in_X2 : INT;
END_VAR
VAR_IN_OUT
	Xus_TN_SCREEN : us_TN_SCREEN;
END_VAR

IF Xus_TN_SCREEN.bya_BACKUP[0] > BYTE#00 THEN

	(* Parameter auslesen *)
	in_X1 := BYTE_TO_INT(Xus_TN_SCREEN.bya_BACKUP[1]);
	in_Y1 := BYTE_TO_INT(Xus_TN_SCREEN.bya_BACKUP[2]);
	in_X2 := BYTE_TO_INT(Xus_TN_SCREEN.bya_BACKUP[3]);
	in_Y2 := BYTE_TO_INT(Xus_TN_SCREEN.bya_BACKUP[4]);

	IF TN_SC_XY2_ERROR(in_X1,in_Y1,in_X2,in_Y2) THEN RETURN; END_IF;
	in_Offset_2 := 5;

	(* CHAR und COLOR von BUFFER wiederherstellen *)
	FOR in_Y := in_Y1 TO in_Y2 DO

		Xus_TN_SCREEN.bya_Line_Update[in_Y] := TRUE; (* Zeile zum Updaten freigeben *)
		in_Offset_1 := (in_Y * 80) + in_X1;

		FOR in_X := in_X1 TO in_X2 DO

			Xus_TN_SCREEN.bya_CHAR[in_Offset_1] := Xus_TN_SCREEN.bya_BACKUP[in_Offset_2];
			in_Offset_2 := in_Offset_2 + INT#01;

			Xus_TN_SCREEN.bya_COLOR[in_Offset_1] := Xus_TN_SCREEN.bya_BACKUP[in_Offset_2];
			in_Offset_2 := in_Offset_2 + INT#01;
			in_Offset_1 := in_Offset_1 + INT#01;

		END_FOR;
	END_FOR;

	(* Daten als ungültig markieren *)
	Xus_TN_SCREEN.bya_BACKUP[0] := BYTE#00;
END_IF;
END_FUNCTION_BLOCK

FUNCTION_BLOCK TN_SC_AREA_SAVE
VAR
	in_Offset_1 : INT;
	in_Offset_2 : INT;
	in_Y : INT;
	in_X : INT;
END_VAR
VAR_INPUT
	Iin_Y1 : INT;
	Iin_X1 : INT;
	Iin_Y2 : INT;
	Iin_X2 : INT;
END_VAR
VAR_IN_OUT
	Xus_TN_SCREEN : us_TN_SCREEN;
END_VAR

IF TN_SC_XY2_ERROR(Iin_X1,Iin_Y1,Iin_X2,Iin_Y2) THEN RETURN; END_IF;

(* Parameter ablegen *)
Xus_TN_SCREEN.bya_BACKUP[0] := BYTE#1;
Xus_TN_SCREEN.bya_BACKUP[1] := INT_TO_BYTE(Iin_X1);
Xus_TN_SCREEN.bya_BACKUP[2] := INT_TO_BYTE(Iin_Y1);
Xus_TN_SCREEN.bya_BACKUP[3] := INT_TO_BYTE(Iin_X2);
Xus_TN_SCREEN.bya_BACKUP[4] := INT_TO_BYTE(Iin_Y2);

in_Offset_2 := 5;
(* CHAR und COLOR in BUFFER sichern *)
FOR in_Y := Iin_Y1 TO Iin_Y2 DO

	in_Offset_1 := (in_Y * 80) + Iin_X1;
	FOR in_X := Iin_X1 TO Iin_X2 DO
		Xus_TN_SCREEN.bya_BACKUP[in_Offset_2] := Xus_TN_SCREEN.bya_CHAR[in_Offset_1];
		in_Offset_2 := in_Offset_2 + INT#01;
		Xus_TN_SCREEN.bya_BACKUP[in_Offset_2] := Xus_TN_SCREEN.bya_COLOR[in_Offset_1];
		in_Offset_2 := in_Offset_2 + INT#01;
		in_Offset_1 := in_Offset_1 + INT#01;
	END_FOR;
END_FOR;
END_FUNCTION_BLOCK

FUNCTION_BLOCK TN_SC_BOX
VAR
	FB_TN_SC_FILL : TN_SC_FILL;
	by_BorderChar_L_T : BYTE;
	by_BorderChar_T : BYTE;
	by_BorderChar_B : BYTE;
	by_BorderChar_R_T : BYTE;
	by_BorderChar_L : BYTE;
	by_BorderChar_R : BYTE;
	by_BorderChar_L_B : BYTE;
	by_BorderChar_R_B : BYTE;
	in_Y : INT;
	in_X : INT;
	in_Border_Offset : INT;
	in_Offset_1 : INT;
	in_Offset_2 : INT;
END_VAR
VAR_INPUT
	Iin_Y1 : INT;
	Iin_X1 : INT;
	Iin_Y2 : INT;
	Iin_X2 : INT;
	Iby_FILL : BYTE;
	Iby_ATTR : BYTE;
	Iin_BORDER : INT;
END_VAR
VAR_IN_OUT
	Xus_TN_SCREEN : us_TN_SCREEN;
END_VAR

IF TN_SC_XY2_ERROR(Iin_X1,Iin_Y1,Iin_X2,Iin_Y2) THEN RETURN; END_IF;

(* Bordertype bestimmen *)
CASE Iin_Border OF
0:
	in_Border_Offset := 0;
1:
	by_BorderChar_L_T := BYTE#218; (* links oben *)
	by_BorderChar_T := BYTE#196; (* oben *)
	by_BorderChar_R_T := BYTE#191; (* rechts oben *)
	by_BorderChar_L := BYTE#179; (* links *)
	by_BorderChar_R := BYTE#179; (* rechts *)
	by_BorderChar_B := BYTE#196; (* unten *)
	by_BorderChar_L_B := BYTE#217; (* links unten *)
	by_BorderChar_R_B := BYTE#192; (* rechts unten *)
	in_Border_Offset := 1;
 2:
	by_BorderChar_L_T := BYTE#201;
	by_BorderChar_T := BYTE#205;
	by_BorderChar_R_T := BYTE#187;
	by_BorderChar_L := BYTE#186;
	by_BorderChar_R := BYTE#186;
	by_BorderChar_B := BYTE#205;
	by_BorderChar_L_B := BYTE#188;
	by_BorderChar_R_B := BYTE#200;
	in_Border_Offset := 1;
ELSE
	by_BorderChar_L_T := BYTE#32;
	by_BorderChar_T := BYTE#32;
	by_BorderChar_R_T := BYTE#32;
	by_BorderChar_L := BYTE#32;
	by_BorderChar_R := BYTE#32;
	by_BorderChar_B := BYTE#32;
	by_BorderChar_L_B := BYTE#32;
	by_BorderChar_R_B := BYTE#32;
	in_Border_Offset := 1;

END_CASE;

IF Iby_FILL > BYTE#0 THEN (* FILL Zeichen vorhanden ? -> Box zeichnen *)

	(* Fill-Function um eine Zeichenreihe kleiner zeichnen *)
	FB_TN_SC_FILL(	Iin_Y1 := Iin_Y1 + in_Border_Offset,
					Iin_X1 := Iin_X1 + in_Border_Offset,
					Iin_Y2 := Iin_Y2 - in_Border_Offset,
					Iin_X2 := Iin_X2 - in_Border_Offset,
					Iby_CHAR := Iby_FILL,
					Iby_Attr := Iby_ATTR,
					Xus_TN_SCREEN := Xus_TN_SCREEN);
END_IF;

IF Iin_BORDER = 0 THEN RETURN; END_IF;

(* linken und rechten Rand ausgeben *)

in_Offset_1 := (Iin_Y1 * 80) + Iin_X1;
in_Offset_2 := (Iin_Y1 * 80) + Iin_X2;

FOR in_Y := Iin_Y1 TO Iin_Y2 DO

	(* Zeile zum Updaten freigeben *)
	Xus_TN_SCREEN.bya_Line_Update[in_Y] := TRUE;

	Xus_TN_SCREEN.bya_CHAR[in_Offset_1] := by_BorderChar_L;
	Xus_TN_SCREEN.bya_COLOR[in_Offset_1] := Iby_Attr;

	Xus_TN_SCREEN.bya_CHAR[in_Offset_2] := by_BorderChar_R;
	Xus_TN_SCREEN.bya_COLOR[in_Offset_2] := Iby_Attr;

	in_Offset_1 := in_Offset_1 + 80;
	in_Offset_2 := in_Offset_2 + 80;

END_FOR;

(* unteren und oberen Rand ausgeben *)
in_Offset_1 := (Iin_Y1 * 80) + Iin_X1;
in_Offset_2 := (Iin_Y2 * 80) + Iin_X1;

FOR in_X := Iin_X1 TO Iin_X2 DO

	Xus_TN_SCREEN.bya_CHAR[in_Offset_1] := by_BorderChar_T;
	Xus_TN_SCREEN.bya_COLOR[in_Offset_1] := Iby_Attr;

	Xus_TN_SCREEN.bya_CHAR[in_Offset_2] := by_BorderChar_B;
	Xus_TN_SCREEN.bya_COLOR[in_Offset_2] := Iby_Attr;

	in_Offset_1 := in_Offset_1 + INT#1;
	in_Offset_2 := in_Offset_2 + INT#1;

END_FOR;

(* linke obere Ecke ausgeben *)
in_Offset_1 := (Iin_Y1 * 80) + Iin_X1;
Xus_TN_SCREEN.bya_CHAR[in_Offset_1] := by_BorderChar_L_T;
Xus_TN_SCREEN.bya_COLOR[in_Offset_1] := Iby_Attr;

(* rechte obere Ecke ausgeben *)
in_Offset_1 := (Iin_Y1 * 80) + Iin_X2;
Xus_TN_SCREEN.bya_CHAR[in_Offset_1] := by_BorderChar_R_T;
Xus_TN_SCREEN.bya_COLOR[in_Offset_1] := Iby_Attr;

(* linke untere Ecke ausgeben *)
in_Offset_1 := (Iin_Y2 * 80) + Iin_X1;
Xus_TN_SCREEN.bya_CHAR[in_Offset_1] := by_BorderChar_R_B;
Xus_TN_SCREEN.bya_COLOR[in_Offset_1] := Iby_Attr;

(* rechte untere Ecke ausgeben *)
in_Offset_1 := (Iin_Y2 * 80) + Iin_X2;
Xus_TN_SCREEN.bya_CHAR[in_Offset_1] := by_BorderChar_L_B;
Xus_TN_SCREEN.bya_COLOR[in_Offset_1] := Iby_Attr;
END_FUNCTION_BLOCK

FUNCTION_BLOCK TN_SC_FILL
VAR
	in_X : INT;
	in_Y : INT;
	in_Offset : INT;
END_VAR
VAR_INPUT
	Iin_Y1 : INT;
	Iin_X1 : INT;
	Iin_Y2 : INT;
	Iin_X2 : INT;
	Iby_CHAR : BYTE;
	Iby_Attr : BYTE;
END_VAR
VAR_IN_OUT
	Xus_TN_SCREEN : us_TN_SCREEN;
END_VAR

IF TN_SC_XY2_ERROR(Iin_X1,Iin_Y1,Iin_X2,Iin_Y2) THEN RETURN; END_IF;

FOR in_Y := Iin_Y1 TO Iin_Y2 DO
	Xus_TN_SCREEN.bya_Line_Update[in_Y] := TRUE; (* Zeile zum Updaten freigeben *)
	in_Offset := (in_Y * 80) + Iin_X1;
	FOR in_X := Iin_X1 TO Iin_X2 DO
		Xus_TN_SCREEN.bya_CHAR[in_Offset]  := Iby_CHAR; (* Zeichen eintragen *)
		Xus_TN_SCREEN.bya_COLOR[in_Offset] := Iby_Attr; (* Farbe eintragen *)
		in_Offset := in_Offset + 1;
	END_FOR;
END_FOR;
END_FUNCTION_BLOCK

FUNCTION_BLOCK TN_SC_LINE
VAR
	by_Connect_Left_Char : BYTE;
	by_Connect_Right_Char : BYTE;
	by_Connect_Top_Char : BYTE;
	by_Connect_Bottom_Char : BYTE;
	by_Connect_Cruz_Char : BYTE;
	by_Vertikal_Line_Char : BYTE;
	by_Horzontal_Line_Char : BYTE;
	by_old_Char : BYTE;
	in_Offset_1 : INT;
	in_ROW_Index : INT;
	in_COL_Index : INT;
	by_Char : BYTE;
END_VAR
VAR_INPUT
	Iin_X1 : INT;
	Iin_Y1 : INT;
	Iin_X2 : INT;
	Iin_Y2 : INT;
	Iby_ATTR : BYTE;
	Iby_BORDER : BYTE;
END_VAR
VAR_IN_OUT
	Xus_TN_SCREEN : us_TN_SCREEN;
END_VAR

IF TN_SC_XY2_ERROR(Iin_X1,Iin_Y1,Iin_X2,Iin_Y2) THEN RETURN; END_IF;

(* Bordertype bestimmen *)
IF Iby_Border = BYTE#01 THEN (* Single Line *)
	by_Connect_Top_Char := BYTE#16#C2;
	by_Connect_Bottom_Char := BYTE#16#C1;
	by_Connect_Left_Char := BYTE#16#C3;
	by_Connect_Right_Char := BYTE#16#B4;
	by_Horzontal_Line_Char := BYTE#16#C4;
	by_Vertikal_Line_Char := BYTE#16#B3;
	by_Connect_Cruz_Char := BYTE#16#C5;
ELSIF Iby_Border = BYTE#02 THEN	(* Double Linie *)
	by_Connect_Top_Char := BYTE#16#CB;
	by_Connect_Bottom_Char := BYTE#16#CA;
	by_Connect_Left_Char := BYTE#16#CC;
	by_Connect_Right_Char := BYTE#16#B9;
	by_Horzontal_Line_Char := BYTE#16#CD;
	by_Vertikal_Line_Char := BYTE#16#BA;
	by_Connect_Cruz_Char := BYTE#16#CE;
ELSE (* Full Linie *)
	by_Connect_Top_Char := Iby_Border;
	by_Connect_Bottom_Char := Iby_Border;
	by_Connect_Left_Char := Iby_Border;
	by_Connect_Right_Char := Iby_Border;
	by_Horzontal_Line_Char := Iby_Border;
	by_Vertikal_Line_Char := Iby_Border;
	by_Connect_Cruz_Char := Iby_Border;
END_IF;

(* Vertikale Linie zeichnen *)
IF Iin_X1 = Iin_X2 THEN
	in_Offset_1 := (Iin_Y1 * 80) + Iin_X1;
	FOR in_ROW_Index := Iin_Y1 TO Iin_Y2 DO
		by_old_Char := Xus_TN_SCREEN.bya_CHAR[in_Offset_1]; (* bestehendes Zeichen auslesen *)
		by_Char := by_Vertikal_Line_Char; (* Standardzeichen vorbelegen *)
		IF by_old_Char = by_Horzontal_Line_Char THEN (* Schnittpunkt erkannt *)
			IF in_ROW_Index = Iin_Y1 THEN (* Anfang der Linie behandeln *)
				by_Char := by_Connect_Top_Char;
			ELSIF in_ROW_Index = Iin_Y2 THEN (* Ende der Linie behandeln *)
				by_Char := by_Connect_Bottom_Char;
			ELSE (* Kreuzungspunkt behandeln *)
				by_Char := by_Connect_Cruz_Char;
			END_IF;
		END_IF;
		Xus_TN_SCREEN.bya_Line_Update[in_ROW_Index] := TRUE; (* Zeile zum Updaten freigeben *)
		Xus_TN_SCREEN.bya_CHAR[in_Offset_1] := by_Char;
		Xus_TN_SCREEN.bya_COLOR[in_Offset_1] := Iby_Attr;
		in_Offset_1 := in_Offset_1 + 80;
	END_FOR;

ELSIF Iin_Y1 = Iin_Y2 THEN (* Horzontale Linie zeichnen *)
	Xus_TN_SCREEN.bya_Line_Update[Iin_Y1] := TRUE; (* Zeile zum Updaten freigeben *)
	in_Offset_1 := (Iin_Y1 * 80) + Iin_X1;
	FOR in_COL_Index := Iin_X1 TO Iin_X2 DO
		by_old_Char := Xus_TN_SCREEN.bya_CHAR[in_Offset_1]; (* bestehendes Zeichen auslesen *)
		by_Char := by_Horzontal_Line_Char; (* Standardzeichen vorbelegen *)
		IF by_old_Char = by_Vertikal_Line_Char THEN (* Schnittpunkt erkannt *)
			IF in_COL_Index = Iin_X1 THEN (* Anfang der Linie behandeln *)
				by_Char := by_Connect_Left_Char;
			ELSIF in_COL_Index = Iin_X2 THEN (* Ende der Linie behandeln *)
				by_Char := by_Connect_Right_Char;
			ELSE (* Kreuzungspunkt behandeln *)
				by_Char := by_Connect_Cruz_Char;
			END_IF;
		END_IF;
		Xus_TN_SCREEN.bya_CHAR[in_Offset_1] := by_Char;
		Xus_TN_SCREEN.bya_COLOR[in_Offset_1] := Iby_Attr;
		in_Offset_1 := in_Offset_1 + 1;
	END_FOR;
END_IF;
END_FUNCTION_BLOCK

FUNCTION_BLOCK TN_SC_READ_ATTR
VAR
	in_Offset : INT;
END_VAR
VAR_INPUT
	Iin_Y : INT;
	Iin_X : INT;
END_VAR
VAR_OUTPUT
	Oby_ATTR : BYTE;
END_VAR
VAR_IN_OUT
	Xus_TN_SCREEN : us_TN_SCREEN;
END_VAR

IF TN_SC_XY_ERROR(Iin_X,Iin_Y) THEN RETURN; END_IF;
in_Offset := (Iin_Y * 80) + Iin_X;
Oby_ATTR := Xus_TN_SCREEN.bya_COLOR[in_Offset]; (* Attribute auslesen *)
END_FUNCTION_BLOCK

FUNCTION_BLOCK TN_SC_READ_CHAR
VAR
	in_Offset : INT;
END_VAR
VAR_INPUT
	Iin_Y : INT;
	Iin_X : INT;
END_VAR
VAR_OUTPUT
	Oby_CHAR : BYTE;
END_VAR
VAR_IN_OUT
	Xus_TN_SCREEN : us_TN_SCREEN;
END_VAR

IF TN_SC_XY_ERROR(Iin_X,Iin_Y) THEN RETURN; END_IF;
in_Offset := (Iin_Y * 80) + Iin_X;
Oby_CHAR := Xus_TN_SCREEN.bya_CHAR[in_Offset]; (* Charakter auslesen *)
END_FUNCTION_BLOCK

FUNCTION TN_SC_SHADOW_ATTR : BYTE
VAR_INPUT
	Iby_ATTR : BYTE;
END_VAR

(* Background Farbe auf Schwarz ändern      *)
(* und dunkle Fordergrundfarben einschalten *)
TN_SC_SHADOW_ATTR := ((Iby_ATTR AND BYTE#2#11110000) OR BYTE#2#00001000);
END_FUNCTION

// Commented out for beedance: it uses FIX, which is commented out.
// FUNCTION_BLOCK TN_SC_VIEWPORT
// VAR
// 	FB_TN_SC_WRITE : TN_SC_WRITE;
// 	FB_TON : TON;
// END_VAR
// VAR
// 	in_index : INT;
// 	in_Color : INT;
// 	by_Attr : BYTE;
// 	in_count : INT;
// END_VAR
// VAR_IN_OUT
// 	Xus_LOG_VIEWPORT : us_LOG_VIEWPORT;
// 	Xus_LOG_CONTROL : LOG_CONTROL;
// 	Xus_TN_SCREEN : us_TN_SCREEN;
// END_VAR
// VAR_INPUT
// 	Iin_X : INT;
// 	Iin_Y : INT;
// 	Iin_Width : INT;
// 	Idw_ATTR_1 : DWORD;
// 	Idw_ATTR_2 : DWORD;
// 	Iti_TIME : TIME;
// END_VAR
//
// (* LOG-Messages ausgeben *)
//
// IF Xus_LOG_VIEWPORT.UPDATE AND FB_TON.Q THEN (* Update gewünscht und Verzögerungszeit abgelaufen *)
// 	Xus_LOG_VIEWPORT.UPDATE := FALSE;
// 	FOR in_count := 1 TO Xus_LOG_VIEWPORT.COUNT DO (* Alle Viewport-Zeilen abarbeiten *)
// 		in_index := Xus_LOG_VIEWPORT.LINE_ARRAY[in_count];
// 		(* Farbe aus den Option-Parameter auslesen >0,Level,Back,Front< *)
// 		in_Color := DWORD_TO_INT(Xus_LOG_CONTROL.MSG_OPTION[in_index] AND DWORD#2#1111);
//
// 		CASE in_Color OF
// 		0..3: by_Attr := BYTE_OF_DWORD(Idw_ATTR_1,INT_TO_BYTE(in_Color));
// 		4..7: by_Attr := BYTE_OF_DWORD(Idw_ATTR_2,INT_TO_BYTE(in_Color));
// 		ELSE
// 			by_Attr := BYTE_OF_DWORD(Idw_ATTR_1,BYTE#0);
// 		END_CASE;
//
// 		(* Message (Text + Farbe) ausgeben *)
// 		FB_TN_SC_WRITE(	Iin_Y := Iin_Y + in_count - INT#01,
// 						Iin_X := Iin_X,
// 						Iby_ATTR := by_Attr,
// 						Ist_STRING := FIX(str := Xus_LOG_CONTROL.MSG[in_index], L := Iin_Width, C := BYTE#32, M := INT#00), (* String rechts ergänzen bzw. kürzen *)
// 						Xus_TN_SCREEN := Xus_TN_SCREEN);
//
// 	END_FOR;
//
// 	(* Timer stoppen/rücksetzen *)
// 	FB_TON.IN := FALSE;
// 	FB_TON.PT := Iti_TIME;
// 	FB_TON();
//
// END_IF;
//
// (* Update-Zeitverzoegerung *)
// FB_TON.IN := TRUE;
// FB_TON.PT := Iti_TIME;
// FB_TON();
// END_FUNCTION_BLOCK

// Commented out for beedance: it uses CODE, which is commented out.
// FUNCTION_BLOCK TN_SC_WRITE
// VAR
// 	bo_Color : BOOL;
// 	in_Offset : INT;
// 	in_Char_Index : INT;
// 	in_String_Length : INT;
// END_VAR
// VAR_INPUT
// 	Iin_Y : INT;
// 	Iin_X : INT;
// 	Iby_ATTR : BYTE;
// 	Ist_STRING : STRING;
// END_VAR
// VAR_IN_OUT
// 	Xus_TN_SCREEN : us_TN_SCREEN;
// END_VAR
//
// in_String_Length := LEN(Ist_STRING);
// IF TN_SC_XY_ERROR(Iin_X + in_String_Length - 1,Iin_Y) THEN RETURN; END_IF;
// Xus_TN_SCREEN.bya_Line_Update[Iin_Y] := TRUE; (* Zeile zum Updaten freigeben *)
// in_Offset := (Iin_Y * 80) + Iin_X; (* Offset des ersten Zeichen berechnen *)
// bo_Color := Iby_ATTR <> BYTE#00;
//
// (* Zeichen und Attribute des String kopieren *)
// FOR in_Char_Index := 1 TO in_String_Length DO
// 	IF bo_Color THEN Xus_TN_SCREEN.bya_COLOR[in_Offset] := Iby_ATTR; END_IF;
// 	Xus_TN_SCREEN.bya_CHAR[in_Offset] := CODE(STR:=Ist_STRING,POS:=in_Char_Index);
// 	in_Offset := in_Offset + INT#1;
// END_FOR;
//
// Xus_TN_SCREEN.in_EOS_Offset := in_Offset; (* End of String Offset sichern *)
// END_FUNCTION_BLOCK

FUNCTION_BLOCK TN_SC_WRITE_ATTR
VAR
	in_Offset : INT;
END_VAR
VAR_INPUT
	Iin_Y : INT;
	Iin_X : INT;
	Iby_ATTR : BYTE;
END_VAR
VAR_IN_OUT
	Xus_TN_SCREEN : us_TN_SCREEN;
END_VAR

IF TN_SC_XY_ERROR(Iin_X,Iin_Y) THEN RETURN; END_IF;
in_Offset := (Iin_Y * 80) + Iin_X;
Xus_TN_SCREEN.bya_COLOR[in_Offset] := Iby_ATTR; (* Attribute schreiben *)
END_FUNCTION_BLOCK

// Commented out for beedance: it uses TN_SC_WRITE, which is commented out.
// FUNCTION_BLOCK TN_SC_WRITE_C
// VAR
// 	FB_TN_SC_WRITE : TN_SC_WRITE;
// END_VAR
// VAR_INPUT
// 	Iin_Y : INT;
// 	Iin_X : INT;
// 	Iby_ATTR : BYTE;
// 	Ist_STRING : STRING;
// 	Iin_LENGTH : INT;
// 	Iin_OPTION : INT;
// END_VAR
// VAR_IN_OUT
// 	Xus_TN_SCREEN : us_TN_SCREEN;
// END_VAR
//
// (* Text ausgeben *)
// FB_TN_SC_WRITE( Iin_Y := Iin_Y,
// 				Iin_X := Iin_X,
// 				Iby_ATTR := Iby_ATTR,
// 				Ist_STRING := FIX(str:=Ist_STRING,L:=Iin_LENGTH,C:=BYTE#32,M:=Iin_OPTION),
// 				Xus_TN_SCREEN := Xus_TN_SCREEN);
// END_FUNCTION_BLOCK

FUNCTION_BLOCK TN_SC_WRITE_CHAR
VAR
	in_Offset : INT;
END_VAR
VAR_INPUT
	Iin_Y : INT;
	Iin_X : INT;
	Iby_CHAR : BYTE;
END_VAR
VAR_IN_OUT
	Xus_TN_SCREEN : us_TN_SCREEN;
END_VAR

IF TN_SC_XY_ERROR(Iin_X,Iin_Y) THEN RETURN; END_IF;
in_Offset := (Iin_Y * 80) + Iin_X;
Xus_TN_SCREEN.bya_CHAR[in_Offset] := Iby_CHAR; (* Charakter schreiben *)
END_FUNCTION_BLOCK

FUNCTION_BLOCK TN_SC_WRITE_EOS
VAR
	TN_SC_WRITE : TN_SC_WRITE;
END_VAR
VAR_INPUT
	Iby_ATTR : BYTE;
	Ist_STRING : STRING;
END_VAR
VAR_IN_OUT
	Xus_TN_SCREEN : us_TN_SCREEN;
END_VAR

TN_SC_WRITE(Iin_Y := Xus_TN_SCREEN.in_EOS_Offset / 80, (* aktuelle Zeile ausrechnen *)
			Iin_X := Xus_TN_SCREEN.in_EOS_Offset MOD 80, (* aktuelle Spalte ausrechnen *)
			Iby_ATTR := Iby_ATTR,
			Ist_STRING := Ist_STRING,
			Xus_TN_SCREEN := Xus_TN_SCREEN);
END_FUNCTION_BLOCK

FUNCTION TN_SC_XY2_ERROR : BOOL
VAR_INPUT
	X1 : INT;
	Y1 : INT;
	X2 : INT;
	Y2 : INT;
END_VAR

(* min und max werte prüfen *)
TN_SC_XY2_ERROR := Y1 < 0 OR X1 < 0 OR Y2 < 0 OR X2 < 0 OR Y1 > 23 OR X1 > 79 OR Y2 > 23 OR X2 > 79;
END_FUNCTION

FUNCTION TN_SC_XY_ERROR : BOOL
VAR_INPUT
	X : INT;
	Y : INT;
END_VAR

(* min und max werte prüfen *)
TN_SC_XY_ERROR := Y < 0 OR X < 0 OR Y > 23 OR X > 79;
END_FUNCTION

FUNCTION_BLOCK TN_SEND_ROWS
VAR_IN_OUT
	IP_C : IP_C;
	S_BUF : NETWORK_BUFFER;
	Xus_TN_SCREEN : us_TN_SCREEN;
END_VAR
VAR_INPUT
	S_BUF_SIZE : INT;
END_VAR
VAR
	in_Line_Count : INT;(*Zähler um max alle 24 Zeilen zu durchlaufen*)
	in_Col_Count : INT;
	in_Last_Row_Index : INT;
	bo_Break_Loop : BOOL;
	in_Row_Count : INT;
	in_Offset : INT;
	in_Write_Index : INT;
	in_Write_Index_Backup : INT;
	by_Cur_Color : BYTE;
	by_last_Color : BYTE;
	in_Write_Stop : INT;
END_VAR

(* Verbindung vorhanden und kein Datensenden aktiv *)
IF (IP_C.C_STATE < BYTE#127 OR S_BUF.SIZE > UINT#0) THEN
	RETURN; (* nein -> Baustein beenden *)
END_IF;

(* aktuellen Schreibindex laden *)
in_Write_Index := UINT_TO_INT(S_BUF.SIZE) - 1;

(* aktuellen Schreibindex zwischenspeichern *)
in_Write_Index_Backup := in_Write_Index;

(* positive Flanke Connect on *)
IF (IP_C.C_STATE = BYTE#254) OR (Xus_TN_SCREEN.bo_Clear_Screen) THEN

	(* Clear-Screen Meldung rücksetzen *)
	Xus_TN_SCREEN.bo_Clear_Screen := FALSE;

	(* alle Zeilen für Update markieren *)
	FOR in_Line_Count := INT#00 TO INT#23 DO
		Xus_TN_SCREEN.bya_Line_Update[in_Line_Count] := TRUE;
	END_FOR;

	(* ESC [0;30,40m  Reset Attributes + Black,Black *)
	in_Write_Index := in_Write_Index + INT#1;
	S_BUF.BUFFER[in_Write_Index] := BYTE#16#1B; (* ESC *)
	in_Write_Index := in_Write_Index + INT#1;
	S_BUF.BUFFER[in_Write_Index] := BYTE#16#5B; (* [ *)
	in_Write_Index := in_Write_Index + INT#1;
	S_BUF.BUFFER[in_Write_Index] := BYTE#16#30; (* 0 *)
	in_Write_Index := in_Write_Index + INT#1;
	S_BUF.BUFFER[in_Write_Index] := BYTE#16#3B; (* ; *)
	in_Write_Index := in_Write_Index + INT#1;
	S_BUF.BUFFER[in_Write_Index] := BYTE#16#33; (* 3 *)

	(* Einerstelle Farbe Foreground ausgeben *)
	in_Write_Index := in_Write_Index + INT#1;
	S_BUF.BUFFER[in_Write_Index] := (SHR(Xus_TN_SCREEN.by_Clear_Screen_Attr,4) OR BYTE#16#30);

	in_Write_Index := in_Write_Index + INT#1;
	S_BUF.BUFFER[in_Write_Index] := BYTE#16#3B; (* ; *)
	in_Write_Index := in_Write_Index + INT#1;
	S_BUF.BUFFER[in_Write_Index] := BYTE#16#34; (* 4 *)

	(* Einerstelle Farbe Background ausgeben *)
	in_Write_Index := in_Write_Index + INT#1;
	S_BUF.BUFFER[in_Write_Index] := ((Xus_TN_SCREEN.by_Clear_Screen_Attr AND BYTE#16#07) OR BYTE#16#30);

	in_Write_Index := in_Write_Index + INT#1;
	S_BUF.BUFFER[in_Write_Index] := BYTE#16#6D; (* m *)

	(* ESC[2J Clear screen and home cursor *)
	in_Write_Index := in_Write_Index + INT#1;
	S_BUF.BUFFER[in_Write_Index] := BYTE#16#1B; (* ESC *)
	in_Write_Index := in_Write_Index + INT#1;
	S_BUF.BUFFER[in_Write_Index] := BYTE#16#5B; (* [ *)
	in_Write_Index := in_Write_Index + INT#1;
	S_BUF.BUFFER[in_Write_Index] := BYTE#16#32; (* 2 *)
	in_Write_Index := in_Write_Index + INT#1;
	S_BUF.BUFFER[in_Write_Index] := BYTE#16#4A; (* J *)

	(* ESC [?7l Off *)
	in_Write_Index := in_Write_Index + INT#1;
	S_BUF.BUFFER[in_Write_Index] := BYTE#16#1B; (* ESC *)
	in_Write_Index := in_Write_Index + INT#1;
	S_BUF.BUFFER[in_Write_Index] := BYTE#16#5B; (* [ *)
	in_Write_Index := in_Write_Index + INT#1;
	S_BUF.BUFFER[in_Write_Index] := BYTE#16#3F; (* ? *)
	in_Write_Index := in_Write_Index + INT#1;
	S_BUF.BUFFER[in_Write_Index] := BYTE#16#37; (* 7 *)
	in_Write_Index := in_Write_Index + INT#1;
	S_BUF.BUFFER[in_Write_Index] := BYTE#16#6C; (* l *)

END_IF;

in_Last_Row_Index := INT#0;
bo_Break_Loop := FALSE;
in_Write_Stop := S_BUF_SIZE - 20;

(* alle Zeilen durchlaufen *)
FOR in_Line_Count := 0 TO 23 DO

	in_Offset := in_Row_Count * INT#80;

	(* prüfen ob Update einer Zeile notwendig ist bzw. nach Reconnect *)
	IF (Xus_TN_SCREEN.bya_Line_Update[in_Row_Count] = TRUE) THEN

		(* Schreib-Cursor positionieren *)
		in_Write_Index := in_Write_Index + INT#1;
		S_BUF.BUFFER[in_Write_Index] := BYTE#16#1B; (* ESC *)
		in_Write_Index := in_Write_Index + INT#1;
		S_BUF.BUFFER[in_Write_Index] := BYTE#16#5B; (* [ *)

		(* Zehnerstelle Zeilennummer ausgeben *)
		in_Write_Index := in_Write_Index + INT#1;
		S_BUF.BUFFER[in_Write_Index] :=
		SHR(INT_TO_BCDC(in_Row_Count + INT#1),INT#4) OR BYTE#16#30;

		(* Einerstelle Zeilennummer ausgeben *)
		in_Write_Index := in_Write_Index + INT#1;
		S_BUF.BUFFER[in_Write_Index] :=
		(INT_TO_BCDC(in_Row_Count + INT#1) AND BYTE#16#0F) OR BYTE#16#30;

		in_Write_Index := in_Write_Index + INT#1;
		S_BUF.BUFFER[in_Write_Index] := BYTE#16#3B; (* ; *)
		in_Write_Index := in_Write_Index + INT#1;
		S_BUF.BUFFER[in_Write_Index] := BYTE#16#31; (* 1 *)
		in_Write_Index := in_Write_Index + INT#1;
		S_BUF.BUFFER[in_Write_Index] := BYTE#16#48; (* H *)

		(* alle Spalten einer Zeile durchlaufen *)
		FOR in_Col_Count := 0 TO 79 DO

			(* aktuelle Farbe bestimmen *)
			by_Cur_Color := Xus_TN_SCREEN.bya_COLOR[in_Offset];
			IF (by_Cur_Color <> by_last_Color) OR (in_Col_Count = INT#00) THEN

				(* Farbeinstellung: ANSI-Sequenz ESC[X;Y;Zm ausgeben *)
				in_Write_Index := in_Write_Index + INT#1;
				S_BUF.BUFFER[in_Write_Index] := BYTE#16#1B; (* ESC *)

				in_Write_Index := in_Write_Index + INT#1;
				S_BUF.BUFFER[in_Write_Index] := BYTE#16#5B; (* [ *)

				(* Farbeinstellung: dunkel oder Hell und blinken bestimmen *)

					IF (((by_Cur_Color AND BYTE#2#10001000) XOR (by_last_Color AND BYTE#2#10001000)) <> BYTE#00) OR (in_Col_Count = 0) THEN

						in_Write_Index := in_Write_Index + INT#1;
						S_BUF.BUFFER[in_Write_Index] := BYTE#16#30; (* 0 *)
						in_Write_Index := in_Write_Index + INT#1;
						S_BUF.BUFFER[in_Write_Index] := BYTE#16#3B; (* ; *)

						(* keine dunklen Farben gewünscht -> dann Bold & Bright *)
						IF (by_Cur_Color AND BYTE#2#00001000) = BYTE#2#00000000 THEN

							(* auf Bold & Btight Farben umstellen *)
							in_Write_Index := in_Write_Index + INT#1;
							S_BUF.BUFFER[in_Write_Index] := BYTE#16#31; (* 1 *)
							in_Write_Index := in_Write_Index + INT#1;
							S_BUF.BUFFER[in_Write_Index] := BYTE#16#3B; (* ; *)

						END_IF;

						(* blinkenden Farben gewünscht *)
						IF (by_Cur_Color AND BYTE#2#10000000) = BYTE#2#10000000 THEN

							(* auf Bold & Bright Farben umstellen *)
							in_Write_Index := in_Write_Index + INT#1;
							S_BUF.BUFFER[in_Write_Index] := BYTE#16#35; (* 5 *)
							in_Write_Index := in_Write_Index + INT#1;
							S_BUF.BUFFER[in_Write_Index] := BYTE#16#3B; (* ; *)

						END_IF;

					END_IF;

					(* Zehnerstelle Farbe Foreground ausgeben *)
					in_Write_Index := in_Write_Index + INT#1;
					S_BUF.BUFFER[in_Write_Index] := BYTE#16#33; (* 3 *)

					(* Einerstelle Farbe Foreground ausgeben *)
					in_Write_Index := in_Write_Index + INT#1;
					S_BUF.BUFFER[in_Write_Index] := ((SHR(by_Cur_Color,4) AND BYTE#2#00000111) OR BYTE#16#30);

					in_Write_Index := in_Write_Index + INT#1;
					S_BUF.BUFFER[in_Write_Index] := BYTE#16#3B; (* ; *)

					(* Zehnerstelle Farbe Background ausgeben *)
					in_Write_Index := in_Write_Index + INT#1;
					S_BUF.BUFFER[in_Write_Index] := BYTE#16#34; (* 4 *)

					(* Einerstelle Farbe Background ausgeben *)
					in_Write_Index := in_Write_Index + INT#1;
					S_BUF.BUFFER[in_Write_Index] := ((by_Cur_Color AND BYTE#2#00000111) OR BYTE#16#30);

					in_Write_Index := in_Write_Index + INT#1;
					S_BUF.BUFFER[in_Write_Index] := BYTE#16#6D; (* m *)

					(* neue Farbe als letzt verwendete speichern *)
					by_last_Color := by_Cur_Color;

				END_IF;

				(* Buffer Ende vorzeitig erreicht -> Ende *)
				IF (in_Write_Index > in_Write_Stop) THEN

					bo_Break_Loop := TRUE;
					EXIT;

				END_IF;

				(* ein TEXT-Zeichen von Screenbuffer in den Sendebuffer übertragen *)
				in_Write_Index := in_Write_Index + INT#1;
				S_BUF.BUFFER[in_Write_Index] := Xus_TN_SCREEN.bya_CHAR[in_Offset];

				(* nächste Spalte anwählen *)
				in_Offset := in_Offset + INT#01;
			END_FOR;

			IF (bo_Break_Loop = TRUE) THEN;

				(* Buffer Ende vorzeitig erreicht -> nur bis zur letzten kompletten Zeile uebertragen *)
				in_Write_Index := in_Last_Row_Index;

				EXIT;
			END_IF;

			(* Buffer ist noch nicht voll -> neue Zeile ubernehmen *)
			in_Last_Row_Index := in_Write_Index;
			Xus_TN_SCREEN.bya_Line_Update[in_Row_Count] := FALSE;

		END_IF;

		(* naechste Zeile adressieren *)
		in_Row_Count := in_Row_Count + INT#01;

		(* ab letzter Zeile wieder von vorne beginnen *)
		IF (in_Row_Count > INT#23) THEN
			in_Row_Count := INT#00;
		END_IF;
		(*-----------------------------------------------*)

	END_FOR;

	(* wenn in einen Update-Zyklus alle Zeilen auf einmal geschafft wurden *)
	(* wird der Row_Count auf ersten Zeile gestellt *)
	(* soll das hässliche Grafikflackern verhindern *)
	(* ansonsten wird bei der letzen Zeile weitergemacht *)
	IF (bo_Break_Loop = FALSE) THEN
		in_Row_Count := INT#00;
	END_IF;

	(* Edit-Cursor positionieren *)
	IF (in_Write_Index <> in_Write_Index_Backup) THEN

		in_Write_Index := in_Write_Index + INT#1;
		S_BUF.BUFFER[in_Write_Index] := BYTE#16#1B; (* ESC *)
		in_Write_Index := in_Write_Index + INT#1;
		S_BUF.BUFFER[in_Write_Index] := BYTE#16#5B; (* [ *)

		(* Zehnerstelle Zeilennummer ausgeben *)
		in_Write_Index := in_Write_Index + INT#1;
		S_BUF.BUFFER[in_Write_Index] := SHR(INT_TO_BCDC(Xus_TN_SCREEN.in_Cursor_Y + 1),INT#4) OR BYTE#16#30;

		(* Einerstelle Zeilennummer ausgeben *)
		in_Write_Index := in_Write_Index + INT#1;
		S_BUF.BUFFER[in_Write_Index] := (INT_TO_BCDC(Xus_TN_SCREEN.in_Cursor_Y + 1) AND BYTE#16#0F) OR BYTE#16#30;

		in_Write_Index := in_Write_Index + INT#1;
		S_BUF.BUFFER[in_Write_Index] := BYTE#16#3B; (* ; *)

		(* Zehnerstelle Spaltenummer ausgeben *)
		in_Write_Index := in_Write_Index + INT#1;
		S_BUF.BUFFER[in_Write_Index] := SHR(INT_TO_BCDC(Xus_TN_SCREEN.in_Cursor_X + 1),INT#4) OR BYTE#16#30;

		(* Einerstelle Spaltennummer ausgeben *)
		in_Write_Index := in_Write_Index + INT#1;
		S_BUF.BUFFER[in_Write_Index] := (INT_TO_BCDC(Xus_TN_SCREEN.in_Cursor_X + 1) AND BYTE#16#0F) OR BYTE#16#30;

		in_Write_Index := in_Write_Index + INT#1;
		S_BUF.BUFFER[in_Write_Index] := BYTE#16#48; (* H *)

END_IF;

(* aktuellen Schreibindex speichern -> Senden anstossen *)
S_BUF.SIZE := INT_TO_UINT(in_Write_Index + 1);
END_FUNCTION_BLOCK

// Commented out for beedance: it uses POINTER TO or ADR, which IEC 61131-3 does not have.
// FUNCTION_BLOCK UNI_CIRCULAR_BUFFER
// VAR_IN_OUT
// 	DATA : UNI_CIRCULAR_BUFFER_DATA;
// END_VAR
// VAR_TEMP
// 	tmp_dw : DWORD;
// 	pTmp : POINTER TO BYTE;
// 	n : INT;
// 	n1 : INT;
// 	n2 : INT;
// 	x: BYTE;
// 	buf_totalsize : UINT;
// END_VAR
// VAR CONSTANT
// 	HeaderSize : INT := 4;
// END_VAR
// VAR
// 	cnt : UINT;
// 	mode_last : INT;
//
// 	(*LOG_MSG : LOG_MSG;
// 	_debug_enable : BOOL := FALSE;*)
// END_VAR
//
// CASE DATA.D_MODE OF
//
// 01:	x := WORD_TO_BYTE(DATA.D_HEAD); (* nur rechtes byte auswerten *)
// 	CASE x OF
// 	01:	cnt := LEN(DATA.D_STRING); (* String verarbeiten *)
// 		pTmp := ADR(DATA.D_STRING);
// 	02:	cnt := 4; (* Real verarbeiten *)
// 		pTmp := ADR(DATA.D_REAL);
// 	03:	cnt := 4; (* DWORD verarbeiten *)
// 		pTmp := ADR(DATA.D_DWORD);
// 	ELSE
// 		cnt := 0;
// 	END_CASE;
//
// 	DATA.BUF_DATA_CNT := DATA.BUF_DATA_CNT + UDINT#1;
//
// 	(* ------ Daten in buffer eintragen ------ *)
// 	buf_totalsize := SIZEOF(DATA.BUF);
//
// 	IF (cnt + HeaderSize) > (buf_totalsize - DATA.BUF_SIZE) THEN (* genug Speicher frei ? *)
// 		DATA.BUF_DATA_LOST := DATA.BUF_DATA_LOST + UDINT#1;
// 		RETURN;
// 	END_IF;
//
// 	DATA.D_SIZE := cnt;
//
// 	mode_last := DATA.D_MODE;
// 	tmp_dw := SHL(WORD_TO_DWORD(DATA.D_HEAD),16) OR UINT_TO_DWORD(cnt);
//
// 	(* Header in Buffer eintragen *)
// 	n1 := 0;
// 	REPEAT
// 		n2 := MIN(HeaderSize - n1, buf_totalsize - DATA._Last);
// 		FOR n := 1 TO n2 DO
// 			tmp_dw := ROL(tmp_dw,8);
// 			data.BUF[DATA._Last] := DWORD_TO_BYTE(tmp_dw);
// 			DATA._Last := DATA._Last + 1;
// 		END_FOR;
// 		IF DATA._Last >= buf_totalsize THEN
// 			DATA._Last := 0;
// 		END_IF
// 		n1 := n1 + n2;
// 	UNTIL n1 >= HeaderSize
// 	END_REPEAT;
//
// 	(* Daten in Buffer eintragen *)
// 	n1 := 0;
// 	REPEAT
// 		n2 := MIN(cnt - n1, buf_totalsize - DATA._Last);
// 		FOR n := 1 TO n2 DO
// 			data.BUF[DATA._Last] := pTmp^;
// 			pTmp := pTmp + 1;
// 			DATA._Last := DATA._Last + 1;
// 		END_FOR;
// 		IF DATA._Last >= buf_totalsize THEN
// 			DATA._Last := 0;
// 		END_IF
// 		n1 := n1 + n2;
// 	UNTIL n1 >= cnt
// 	END_REPEAT;
//
// 	DATA.BUF_SIZE := DATA.BUF_SIZE + cnt + HeaderSize;
// 	DATA.BUF_COUNT := DATA.BUF_COUNT + 1;
// 	DATA.BUF_USED := UINT_TO_USINT(100 * DATA.BUF_SIZE / buf_totalsize); (* benützer Speicher in % *)
// 	DATA.D_MODE := 0;
//
// 	(*####################  DEBUG-MESSAGE  ###################################*)
// 	(*IF _debug_enable THEN
// 		LOG_CL.NEW_MSG := 'RP: ADD /HEAD ~1 / SIZE ~2 / CNT ~3 / >~4<';
// 		LOG_CL.PRINTF[1] := DWORD_TO_STRH(DATA.D_HEAD);
// 		LOG_CL.PRINTF[2] := UINT_TO_STRING(cnt);
// 		LOG_CL.PRINTF[3] := UINT_TO_STRING(DATA.BUF_COUNT);
// 		CASE x OF
// 		01:	LOG_CL.PRINTF[4] := DATA.D_STRING;
// 		02:	LOG_CL.PRINTF[4] := REAL_TO_STRING(DATA.D_REAL);
// 		03:	LOG_CL.PRINTF[4] := DWORD_TO_STRH(DATA.D_DWORD);
// 		ELSE
// 			LOG_CL.PRINTF[4] := '';
// 		END_CASE;
// 		LOG_MSG();
// 	END_IF;*)
// 	(*########################################################################*)
//
// 10..12:	(* ------ Daten aus buffer auslesen und optional löschen ------ *)
// 		(* 10 = nur lesen / 11 = löschen nach lesen / 12 = lesen und löschen *)
// 	IF DATA.D_MODE <> 11 THEN
// 		IF DATA.BUF_COUNT = 0 THEN RETURN; END_IF;
// 		buf_totalsize := SIZEOF(DATA.BUF);
// 		DATA._GetEnd := DATA._First;(* index des ältesten eintrags merken *)
// 		mode_last := DATA.D_MODE;
//
// 		(* Header aus Buffer lesen *)
// 		n1 := 0;
// 		tmp_dw := 0;
// 		REPEAT
// 			n2 := MIN(HeaderSize - n1, buf_totalsize - DATA._GetEnd);
// 			FOR n := 1 TO n2 DO
// 				tmp_dw := ROL(tmp_dw,8) OR BYTE_TO_DWORD(data.BUF[DATA._GetEnd]);
// 				DATA._GetEnd := DATA._GetEnd + 1;
// 			END_FOR;
// 			IF DATA._GetEnd >= buf_totalsize THEN
// 				DATA._GetEnd := 0;
// 			END_IF
// 			n1 := n1 + n2;
// 		UNTIL n1 >= HeaderSize
// 		END_REPEAT;
//
// 		DATA._GetStart := DATA._GetEnd;
// 		cnt := DWORD_TO_UINT(tmp_dw AND 16#0000_FFFF);
// 		DATA.D_SIZE := cnt;
// 		DATA.D_HEAD := DWORD_TO_WORD(SHR(tmp_dw,16));
//
// 		x := WORD_TO_BYTE(DATA.D_HEAD); (* nur rechtes byte auswerten *)
// 		CASE x OF
// 		01:	pTmp := ADR(DATA.D_STRING); (* String verarbeiten *)
// 		02:	pTmp := ADR(DATA.D_REAL); (* Real verarbeiten *)
// 		03:	pTmp := ADR(DATA.D_DWORD); (* DWORD verarbeiten *)
// 		END_CASE;
//
// 		(* Daten aus Buffer lesen *)
// 		n1 := 0;
// 		REPEAT
// 			n2 := MIN(cnt - n1, buf_totalsize - DATA._GetEnd);
// 			FOR n := 1 TO n2 DO
// 				pTmp^ := data.BUF[DATA._GetEnd];
// 				pTmp := pTmp + 1;
// 				DATA._GetEnd := DATA._GetEnd + 1;
// 			END_FOR;
// 			IF DATA._GetEnd >= buf_totalsize THEN
// 				DATA._GetEnd := 0;
// 			END_IF
// 			n1 := n1 + n2;
// 		UNTIL n1 >= cnt
// 		END_REPEAT;
// 		IF x = 1 THEN
// 			pTmp^ := 0; (* String terminieren *)
// 		END_IF;
// 		DATA.D_MODE := 0;
//
// 		(*####################  DEBUG-MESSAGE  ###################################*)
// 		(*IF _debug_enable THEN
// 			LOG_CL.NEW_MSG := 'RP: READ /HEAD ~1 / SIZE ~2 / CNT ~3 / >~4<';
// 			LOG_CL.PRINTF[1] := DWORD_TO_STRH(DATA.D_HEAD);
// 			LOG_CL.PRINTF[2] := UINT_TO_STRING(cnt);
// 			LOG_CL.PRINTF[3] := UINT_TO_STRING(DATA.BUF_COUNT);
// 			CASE x OF
// 			01:	LOG_CL.PRINTF[4] := DATA.D_STRING;
// 			02:	LOG_CL.PRINTF[4] := REAL_TO_STRING(DATA.D_REAL);
// 			03:	LOG_CL.PRINTF[4] := DWORD_TO_STRH(DATA.D_DWORD);
// 			ELSE
// 				LOG_CL.PRINTF[4] := '';
// 			END_CASE;
// 			LOG_MSG();
// 		END_IF;*)
// 		(*########################################################################*)
// 	END_IF;
//
// 	IF (mode_last = 10 AND DATA.D_MODE = 11) OR (mode_last = 12 AND DATA.D_MODE = 0) THEN (* löschen nur direkt nach lesen möglich *)
// 		mode_last := DATA.D_MODE;
// 		DATA.BUF_SIZE := DATA.BUF_SIZE - cnt - HeaderSize;
// 		DATA.BUF_COUNT := DATA.BUF_COUNT - 1;
// 		DATA._First := DATA._GetEnd;
// 		DATA.BUF_USED := UINT_TO_USINT(100 * DATA.BUF_SIZE / SIZEOF(DATA.BUF)); (* benützer Speicher in % *)
// 		DATA.D_MODE := 0;
//
// 		(*####################  DEBUG-MESSAGE  ###################################*)
// 		(*IF _debug_enable THEN
// 			LOG_CL.NEW_MSG := 'RP: DEL /HEAD ~1 / SIZE ~2 / CNT ~3 / >~4<';
// 			LOG_CL.PRINTF[1] := DWORD_TO_STRH(DATA.D_HEAD);
// 			LOG_CL.PRINTF[2] := UINT_TO_STRING(cnt);
// 			LOG_CL.PRINTF[3] := UINT_TO_STRING(DATA.BUF_COUNT);
// 			CASE x OF
// 			01:	LOG_CL.PRINTF[4] := DATA.D_STRING;
// 			02:	LOG_CL.PRINTF[4] := REAL_TO_STRING(DATA.D_REAL);
// 			03:	LOG_CL.PRINTF[4] := DWORD_TO_STRH(DATA.D_DWORD);
// 			ELSE
// 				LOG_CL.PRINTF[4] := '';
// 			END_CASE;
// 			LOG_MSG();
// 		END_IF;*)
// 		(*########################################################################*)
// 	END_IF;
//
// 99:	(* Buffer reset - alles löschen *)
// 	DATA._First := 0;
// 	DATA._Last := 0;
// 	DATA._GetStart := 0;
// 	DATA._GetEnd := 0;
// 	DATA.BUF_COUNT := 0;
// 	DATA.BUF_SIZE := 0;
// 	DATA.BUF_USED := 0;
// 	DATA.D_STRING := '';
// 	DATA.D_DWORD := 0;
// 	DATA.D_REAL := 0.0;
// 	DATA.D_HEAD := 0;
// 	DATA.D_MODE := 0;
// 	DATA.D_SIZE := 0;
// 	mode_last := 0;
// END_CASE;
//
// (* höchsten Auslastungswert speichern *)
// IF DATA.BUF_USED > DATA.BUF_USED_MAX THEN
// 	DATA.BUF_USED_MAX := DATA.BUF_USED;
// END_IF;
// END_FUNCTION_BLOCK

// Commented out for beedance: it uses CHR_TO_STRING, which is commented out.
// FUNCTION URL_DECODE : STRING(STRING_LENGTH)
// VAR_INPUT
// 	IN : STRING(STRING_LENGTH);
// END_VAR
// VAR
// 	pos : INT;
// 	seq : STRING(3);
// 	new : STRING(1);
// END_VAR
//
// URL_DECODE := IN;
// pos := FIND(URL_DECODE,'%');
// WHILE pos > 0 DO
// 	seq := MID(URL_DECODE,2,pos + 1);
// 	new := CHR_TO_STRING(DWORD_TO_BYTE(HEX_TO_DWORD(seq)));
// 	URL_DECODE := REPLACE(URL_DECODE, new, 3, pos);
// 	pos := FIND(URL_DECODE,'%');
// END_WHILE;
// END_FUNCTION

// Commented out for beedance: it uses POINTER TO or ADR, which IEC 61131-3 does not have.
// FUNCTION URL_ENCODE : STRING(STRING_LENGTH)
// VAR_INPUT
// 	IN : STRING(STRING_LENGTH);
// END_VAR
// VAR
// 	pt_in : POINTER TO ARRAY[1..255] OF BYTE;
// 	pt_out : POINTER TO ARRAY[1..256] OF BYTE;
// 	pos_in : INT;
// 	pos_out : INT;
// 	stop : INT;
// 	tb : BYTE;
// END_VAR
//
// pt_in  := ADR(in);
// pt_out := ADR(URL_ENCODE);
//
// (* scan the input string and convert unallowed characters *)
// pos_in := 1;
// stop := LEN(in);
// FOR pos_out := 1 TO 250 DO
// 	IF pos_in > stop THEN
// 		EXIT;
// 	ELSIF IS_URLCHR(pt_in^[pos_in]) THEN
// 		pt_out^[pos_out] := pt_in^[pos_in];
// 		(* increment in by 1 *)
// 		pos_in := pos_in + 1;
// 	ELSE
// 		(* cannot fit 3 digits, exit *)
// 		IF pos_out > 248 THEN EXIT; END_IF;
// 		(* invalid character that needs to be converted *)
// 		pt_out^[pos_out] := 37;    (* start with % sign *)
// 		pos_out := pos_out + 1;
// 		(* need to add the two hex digits *)
// 		tb := SHR(pt_in^[pos_in],4);
// 		IF tb > 9 THEN
// 			pt_out^[pos_out] := tb + 55;
// 		ELSE
// 			pt_out^[pos_out] := tb + 48;
// 		END_IF;
// 		pos_out := pos_out + 1;
// 		tb := pt_in^[pos_in] AND 16#0F;
// 		IF tb > 9 THEN
// 			pt_out^[pos_out] := tb + 55;
// 		ELSE
// 			pt_out^[pos_out] := tb + 48;
// 		END_IF;
// 		(* increment in and out because out has to move 3 digits *)
// 		pos_in := pos_in + 1;
// 	END_IF;
// END_FOR;
//
// (* terminate the output string *)
// pt_out^[pos_out] := 0;
// END_FUNCTION

FUNCTION URL_TO_STRING : STRING(STRING_LENGTH)
VAR_INPUT
	IN : URL;
END_VAR

(*

http://hans:geheim@www.example.org:80/demo/example.cgi?land=de&stadt=aa#abschnitt1
|         |         |                  |                                |   |                                    |                                    |
|         |         |                 Host                         |   Pfad                            Query                           Anker
|         |         Passwort                                  Port
|        Benutzer
Protokoll

*)

(* attach protocol *)
IF IN.PROTOCOL <> '' THEN URL_TO_STRING := CONCAT(IN.PROTOCOL,'://'); END_IF;

(* attach user and password *)
IF IN.USER <> '' THEN
	URL_TO_STRING := CONCAT(URL_TO_STRING, IN.USER);
	IF IN.PASSWORD <> '' THEN
		URL_TO_STRING := CONCAT(URL_TO_STRING, ':');
		URL_TO_STRING := CONCAT(URL_TO_STRING, IN.PASSWORD);
	END_IF;
	URL_TO_STRING := CONCAT(URL_TO_STRING, '@');
END_IF;

(* attach domain *)
URL_TO_STRING := CONCAT(URL_TO_STRING, IN.DOMAIN);

(* attach Port *)
IF IN.PORT > 0 THEN
	URL_TO_STRING := CONCAT(URL_TO_STRING, ':');
	URL_TO_STRING := CONCAT(URL_TO_STRING, WORD_TO_STRING(IN.PORT));
END_IF;

(* attach path *)
URL_TO_STRING := CONCAT(URL_TO_STRING, IN.PATH);

(* attach query *)
IF IN.QUERY <> '' THEN
	URL_TO_STRING := CONCAT(URL_TO_STRING, '?');
	URL_TO_STRING := CONCAT(URL_TO_STRING, IN.QUERY);
END_IF;

(* attach anchor *)
IF IN.ANCHOR <> '' THEN
	URL_TO_STRING := CONCAT(URL_TO_STRING, '#');
	URL_TO_STRING := CONCAT(URL_TO_STRING, IN.ANCHOR);
END_IF;
END_FUNCTION

// Commented out for beedance: it uses CSV_PARSER_BUF, which is commented out.
// FUNCTION_BLOCK WORLD_WEATHER
// VAR_IN_OUT
// 	IP_C : IP_C; (* IP_Control Verwaltungsstruktur *)
// 	S_BUF : NETWORK_BUFFER;
// 	R_BUF : NETWORK_BUFFER;
// 	WW : WORLD_WEATHER_DATA;
// END_VAR
// VAR_INPUT
// 	ACTIVATE : BOOL;
// 	LATITUDE : REAL;
// 	LONGITUDE : REAL;
// 	KEY : STRING(30);
// END_VAR
// VAR_OUTPUT
// 	BUSY : BOOL;
// 	DONE : BOOL;
// 	ERROR_C : DWORD;
// 	ERROR_T : BYTE;
// END_VAR
// VAR
// 	URL_DATA : url;
// 	DNS_CLIENT : DNS_CLIENT;
// 	HTTP_GET : HTTP_GET;
// 	CPB : CSV_PARSER_BUF;
// 	last_state : BOOL;
// 	value_int : INT;
// 	value_real : REAL;
// 	v_real : REAL;
// 	state : INT;
// 	url_str : STRING(STRING_LENGTH);
// 	offset : UDINT;
// 	size : INT;
// 	sep : BYTE;
// 	cnt : INT;
// 	day : INT;
// 	idx : INT;
// 	run : BYTE;
// 	result : BYTE;
// 	value : STRING(STRING_LENGTH);
// 	pos : INT;
// END_VAR
//
// CASE state OF
//
// 00:
// 	IF ACTIVATE AND NOT last_state THEN
// 		state := 20;
// 		DONE := FALSE;
// 		BUSY := TRUE;
// 		ERROR_C := DWORD#0;
// 		ERROR_T := BYTE#0;
// 	END_IF;
//
// 20: (* URL for DNS UND HTTP-GET *)
// 	(* Example: http://api.worldweatheronline.com/free/v1/weather.ashx?q=48.21,16.37&format=csv&num_of_days=5&key=xxxxxxxxxxxxxxxxxxxxxx *)
// 	url_str := CONCAT('http://api.worldweatheronline.com/free/v1/weather.ashx?q=',REAL_TO_STRF(LATITUDE,6,D:='.'));
// 	url_str := CONCAT(url_str,',');
// 	url_str := CONCAT(url_str,REAL_TO_STRF(LONGITUDE,6,D:='.'));
// 	url_str := CONCAT(url_str,'&format=csv&num_of_days=5&key=');
// 	url_str := CONCAT(url_str,key);
//
// 	URL_DATA:=STRING_TO_URL(STR:=url_str, DEFAULT_PROTOCOL:='', DEFAULT_PATH:='' );
// 	state := 40;
//
// 40:
// 	IF DNS_CLIENT.DONE THEN
// 		state := 60;
// 	ELSIF (DNS_CLIENT.ERROR > DWORD#00) THEN
// 		(* Fehlerbehandlung *)
// 		ERROR_C := DNS_CLIENT.ERROR;
// 	ERROR_T := BYTE#01;
// 		state   := 100;
// 	END_IF;
//
// 60:
// 	IF HTTP_GET.DONE THEN
// 		sep := 0;
// 		idx := 0;
// 		day := 0;
// 		cnt := 0;
// 		OFFSET := HTTP_GET.BODY_START; (* Start Offset vorgeben *)
// 		size := HTTP_GET.BODY_STOP; (* End Position *)
// 		run := 1; (* Element suchen *)
// 		state := 80;
//
// 	ELSIF (HTTP_GET.ERROR > DWORD#00) THEN
// 		(* Fehlerbehandlung *)
// 		ERROR_C := HTTP_GET.ERROR;
// 		ERROR_T := BYTE#02;
// 		state := 100;
// 	END_IF;
//
// 80:	IF run = 0 THEN (* kein Befehl mehr aktiv ? *)
// 		run := 1; (*  nächstes Element suchen  *)
// 		IF result = 1 OR result = 2 THEN
// 			value_int := 0;
// 			value_real := 0.0;
// 			(* automatische konvertierung in real und int ausführen *)
// 			IF LEN(value) <= 20 THEN
// 				v_real:=FLOAT_TO_REAL(FLT:=value);
// 				IF CHK_REAL(v_real) = 0 THEN (* !!! prüft auf gültigen REAL Wert, ansonsten stürzt Twincat ab !!!!  *)
// 					value_real := v_real;
// 					value_int := REAL_TO_INT(value_real);
// 				END_IF;
// 			END_IF;
// 			cnt := cnt + 1;
//
// 			IF cnt = 1 AND LEFT(value,1) <> '#' THEN
// 				cnt := 0;
// 			END_IF;
//
// 			IF cnt >=8 AND cnt <= 87 THEN
// 				IF cnt > 22 THEN
// 					CASE idx OF
// 					00:	WW.DAY[day].DATE_OF_DAY := value;
// 					01:	WW.DAY[day].TEMP_MAX_C := value_int;
// 					02:	WW.DAY[day].TEMP_MAX_F := value_int;
// 					03:	WW.DAY[day].TEMP_MIN_C := value_int;
// 					04:	WW.DAY[day].TEMP_MIN_F := value_int;
// 					05:	WW.DAY[day].WIND_SPEED_MILES := value_int;
// 					06:	WW.DAY[day].WIND_SPEED_KMPH := value_int;
// 					07:	WW.DAY[day].WIND_DIR_DEGREE := value_int;
// 					08:	WW.DAY[day].WIND_DIR16POINT := value;
// 					09:	WW.DAY[day].WEATHER_CODE := value_int;
// 					10:	pos := FIND(value, '/wsymbol_');
// 						WW.DAY[day].WEATHER_ICON := DEC_TO_INT(MID(value,4,pos+9));
// 					11:	WW.DAY[day].WEATHER_DESC := value;
// 					12:	WW.DAY[day].PRECIPMM := value_real;
// 					END_CASE;
// 					idx := idx + 1;
// 					IF idx > 12 THEN
// 						idx := 0;
// 						day := day + 1;
// 					END_IF;
// 				ELSE
// 					CASE cnt OF
// 					08:	sep :=44; (* ab jetzt mit Trennzeichen arbeiten, *)
// 					09:	WW.CUR.OBSERVATION_TIME := value;
// 					10:	WW.CUR.TEMP_C := value_int;
// 					11:	WW.CUR.WEATHER_CODE := value_int;
// 					12:	pos := FIND(value, '/wsymbol_');
// 						WW.CUR.WEATHER_ICON := DEC_TO_INT(MID(value,4,pos+9));
// 					13:	WW.CUR.WEATHER_DESC := value;
// 					14:	WW.CUR.WIND_SPEED_MILES := value_int;
// 					15:	WW.CUR.WIND_SPEED_KMPH := value_int;
// 					16:	WW.CUR.WIND_DIR_DEGREE := value_int;
// 					17:	WW.CUR.WIND_DIR16POINT := value;
// 					18:	WW.CUR.PRECIPMM := value_real;
// 					19:	WW.CUR.HUMIDITY := value_int;
// 					20:	WW.CUR.VISIBILITY := value_int;
// 					21:	WW.CUR.PRESSURE := value_int;
// 					22:	WW.CUR.CLOUDOVER := value_int;
// 					END_CASE;
// 				END_IF;
// 			END_IF;
// 		ELSIF result = 10 THEN (* nichts mehr gefunden *)
// 			DONE  := TRUE;
// 			run := 0; (* Auswertung beenden *)
// 			state := 100;
// 		END_IF;
// 	END_IF;
//
// 100:
// 	(* UNLOCK HTTP DATA *)
// 	IF (NOT HTTP_GET.DONE) THEN
// 		state := 0;
// 		BUSY := FALSE;
// 		DONE := ERROR_T = BYTE#0;
// 	END_IF;
//
// END_CASE;
//
// (* ---------------- DNS --------------- *)
// DNS_CLIENT(	IP_C:=IP_C,
// 			S_BUF:=S_BUF,
// 			R_BUF:=R_BUF,
// 			DOMAIN:=URL_DATA.DOMAIN,
// 			IP4_DNS:=DWORD#00,
// 			ACTIVATE:=state=40 (* DNS Start *)
// 			);
// (* nicht oder nicht direkt verwendete Parameter *)
// (*	DWORD :=DNS_CLIENT.IP4;
// 	BOOL  :=DNS_CLIENT.DONE;
// 	BYTE  :=DNS_CLIENT.ERROR; *)
// (* -------------------------------------*)
//
// (* ------------- HTTP_GET --------------- *)
// HTTP_GET(	IP_C:=IP_C,
// 			S_BUF:=S_BUF,
// 			R_BUF:=R_BUF,
// 			IP4:=DNS_CLIENT.IP4,
// 			GET:=state=60,
// 			MODE:=BYTE#2, (* HTTP 1.1 mit persistenter Verbindung *)
// 			UNLOCK_BUF:=state=100,
// 			URL_DATA:=URL_DATA
// 			);
//
// (* nicht oder nicht direkt verwendete Parameter *)
// (*	STRING := HTTP_GET.HTTP_STATUS;
// 	UINT :=HTTP_GET.HEADER_START;
// 	UINT :=HTTP_GET.HEADER_STOP;
// 	UINT :=HTTP_GET.BODY_START;
// 	UINT :=HTTP_GET.BODY_STOP;
// 	BOOL :=HTTP_GET.DONE;
// 	BYTE :=HTTP_GET.ERROR;
// *)
// (* -------------------------------------*)
// CPB(SEP:=sep,RUN:=run,OFFSET:=OFFSET,VALUE:=value,PT:=R_BUF,RESULT=>result); (* CSV PARAMETER BUF *)
//
// last_state := ACTIVATE;
// END_FUNCTION_BLOCK

FUNCTION_BLOCK WORLD_WEATHER_DESC_GE
VAR_IN_OUT
	WW : WORLD_WEATHER_DATA;
END_VAR
VAR_INPUT
	ACTIVATE : BOOL;
END_VAR
VAR
	act_last : BOOL;
	x : INT;
	y : INT;
	str : STRING(60);
	i : INT;
END_VAR

IF ACTIVATE AND act_last = FALSE THEN
	i := 0;
	FOR y := 1 TO 12 DO
		CASE y OF
		1,3,5,7,9:		x :=  WW.DAY[i].WEATHER_CODE;
		2,4,6,8,10:	WW.DAY[i].WEATHER_DESC := str;
					i := i + 1;
		11:			x :=  WW.CUR.WEATHER_CODE;
		12:			WW.CUR.WEATHER_DESC := str;
		END_CASE;

		CASE x OF
			113	:	str := 'heiter/sonnig';
			116	:	str := 'stellenweise wolkig';
			119	:	str := 'wolkig';
			122	:	str := 'bewölkt';
			143	:	str := 'Nebel';
			176	:	str := 'stellenweise nahegelegener Regen';
			179	:	str := 'stellenweise nahegelegener Schneefall';
			182	:	str := 'stellenweise nahegelegener Eisregen';
			185	:	str := 'stellenweise gefrierender Niesel';
			200	:	str := 'nahegelegene Sturm';
			227	:	str := 'Schneetreiben';
			230	:	str := 'Schneesturm';
			248	:	str := 'Nebel';
			260	:	str := 'gefrierender Nebel';
			263	:	str := 'stellenweise leichter Nieselregen';
			266	:	str := 'leichter Niesel';
			281	:	str := 'gefrierender Nieselregen';
			284	:	str := 'stark gefrierender Nieselregen';
			293	:	str := 'stellenweise leichter Regen';
			296	:	str := 'leichter Regen';
			299	:	str := 'zeitweise etwas Regen';
			302	:	str := 'mäßiger Regen';
			305	:	str := 'zeitweise etwas starker Regen';
			308	:	str := 'starker Regen';
			311	:	str := 'leichter gefrierender Regen';
			314	:	str := 'mäßiger oder starker Eisregen';
			317	:	str := 'leichter Eisregen';
			320	:	str := 'mäßiger oder starker Eisregen';
			323	:	str := 'stellenweise leichter Schneefall';
			326	:	str := 'leichter Scheefall';
			329	:	str := 'stellenweise moderater Schneefall';
			332	:	str := 'mäßiger Schnee';
			335	:	str := 'stellenweise starker Scheefall';
			338	:	str := 'starker Schneefall';
			350	:	str := 'Hagel';
			353	:	str := 'leichte Regenfälle';
			356	:	str := 'mäßiger oder starker Regenfall';
			359	:	str := 'sintflutartige Regenfälle';
			362	:	str := 'leichter Eisregen';
			365	:	str := 'mäßiger oder starker Eisregen';
			368	:	str := 'leichte Schneeschauer';
			371	:	str := 'mäßiger oder starker Schneefall';
			374	:	str := 'leichter Hagel';
			377	:	str := 'mäßiger oder starker Hagel';
			386	:	str := 'stellenweise leichter Regen in Gewittergebiet';
			389	:	str := 'mäßiger oder starker Regen in Gewittergebiet';
			392	:	str := 'stellenweise leichter Schneefall in Gewittergebiet';
			395	:	str := 'mäßiger oder starker Schnee in Gewittergebiet';
		ELSE
			str := 	'nicht verfügbar';
		END_CASE;
	END_FOR;
END_IF;
act_last := ACTIVATE;
END_FUNCTION_BLOCK

FUNCTION_BLOCK WORLD_WEATHER_ICON_OSCAT
VAR_IN_OUT
	WW : WORLD_WEATHER_DATA;
END_VAR
VAR_INPUT
	ACTIVATE : BOOL;
END_VAR
VAR
	dat : ARRAY[0..41] OF INT := 0,14,12,9,9,0,7,7,0,2,2,3,3,1,0,0,17,4,4,3,3,1,0,0,17,2,2,3,3,1,0,0,17,2,4,3,3,1,0,0,17,0;
	act_last : BOOL;
	x : INT;
	i : INT;
END_VAR

IF ACTIVATE AND act_last = FALSE THEN
	x := LIMIT(0,WW.CUR.WEATHER_ICON,41);
	WW.CUR.WEATHER_ICON := dat[x];
	FOR i := 0 TO 4 DO
		x := LIMIT(0,WW.DAY[i].WEATHER_ICON,41);
		WW.DAY[i].WEATHER_ICON := dat[x];
	END_FOR;
END_IF;
act_last := ACTIVATE;
END_FUNCTION_BLOCK

// Commented out for beedance: it uses POINTER TO or ADR, which IEC 61131-3 does not have.
// FUNCTION_BLOCK XML_READER
// VAR_IN_OUT
// 	CTRL : XML_CONTROL;
// 	BUF : NW_BUF_LONG;
// END_VAR
// VAR
// 	index :	INT;
// 	index2 : INT;
// 	stop : INT;
// 	mode : INT;
// 	command : WORD;
// 	c :	BYTE;
// 	s1 : INT;
// 	e1 : INT;
// 	path_overflow : BOOL;
// 	empty_tag : BOOL;
// 	s_code : STRING(10);
// 	e_code : STRING(10);
// 	watchdog : TON;
//
// 	(*LOG_MSG : LOG_MSG;
// 	_debug_enable : BOOL := TRUE;*)
//
// END_VAR
//
// (*
//
// TYP
// 00 = UNBEKANNT
// 01 = ELEMENT (STANDARD)
// 02 = CLOSE ELEMENT
// 03 = TEXT
// 04 = ATTRIBUTE
// 05 = ELEMENT (PROCESSING INSTRUCTION)
//
// 12 = !CDATA
// 13 = !COMMENT
// 14 = !DTD ELEMENT (Document Type Declarations )
//
// 98 = WATCHDOG
// 99 = ENDE
//
// Bei Typ 02 werden keine Blockdaten ausgegeben !
//
// *)
//
// (* ---------- Init -------------- *)
// IF BIT_OF_DWORD(WORD_TO_DWORD(CTRL.COMMAND),15) THEN
// 	COMMAND := CTRL.COMMAND;
// 	CTRL.COMMAND := WORD#0;
//
// 	index := UINT_TO_INT(CTRL.START_POS);
// 	stop := UINT_TO_INT(CTRL.STOP_POS);
// 	mode := 100;
// 	path_overflow := FALSE;
//
// 	CTRL.TYP := 0;
// 	CTRL.COUNT := UINT#00;
// 	CTRL.LEVEL := UINT#00;
// 	CTRL.ATTRIBUTE := '';
// 	CTRL.ELEMENT := '';
// 	CTRL.PATH := '';
// 	CTRL.VALUE := '';
//
// 	WATCHDOG.PT := CTRL.WATCHDOG;
// END_IF;
//
// (*----------------------------------------------- *)
//
// IF index < 0 THEN RETURN;END_IF;
//
// CTRL.BLOCK1_START := UINT#0;
// CTRL.BLOCK1_STOP := UINT#0;
// CTRL.BLOCK2_START := UINT#0;
// CTRL.BLOCK2_STOP := UINT#0;
//
// WATCHDOG(IN:=FALSE); (* Timer stoppen *)
//
// WHILE (TRUE) DO
//
// 	(* -------------- WATCHDOG ------------------ *)
// 	WATCHDOG(IN:=CTRL.WATCHDOG > T#0s);
// 	IF WATCHDOG.Q THEN
// 		CTRL.TYP := 98;
//     		(*####################  DEBUG-MESSAGE  ###################################*)
//     		(*IF _debug_enable THEN
//       			LOG_CL.NEW_MSG := 'WATCHDOG:';
//       			LOG_MSG();
//     		END_IF;*)
//     		(*########################################################################*)
// 		RETURN;
// 	END_IF;
//
// 	(* -------------- PARSING END ------------------ *)
// 	IF index > stop THEN
// 		CTRL.COUNT := CTRL.COUNT + UINT#1;
// 		CTRL.TYP := 99;
//     		(*####################  DEBUG-MESSAGE  ###################################*)
//     		(*IF _debug_enable THEN
//       			LOG_CL.NEW_MSG := 'EX: #T:~1 #C:~2 #P:~6 #L:~7';
//       			LOG_CL.PRINTF[1] := INT_TO_STRING(CTRL.TYP);
//       			LOG_CL.PRINTF[2] := UINT_TO_STRING(CTRL.COUNT);
//       			LOG_CL.PRINTF[6] := CTRL.PATH;
//       			LOG_CL.PRINTF[7] := UINT_TO_STRING(CTRL.LEVEL);
//       			LOG_MSG();
//     		END_IF;*)
//     		(*########################################################################*)
// 		mode  := 0; (* Schritt ruecksetzen *)
// 		index := 0; (* Abarbeitung stoppen *)
// 		RETURN;
// 	END_IF;
//
// 	CASE mode OF
//
// 	100: (* ---------- ELEMENT SECTION ------------------ *)
// 		(* search begin of element *)
// 		s1 := 0;
// 		e1 := 0;
// 		WHILE (index <= stop) DO
// 			IF BUF[INDEX]=BYTE#60 THEN (* '<' TagBegin *)
// 				index := index + 1;
// 				C := BUF[index];
// 				IF C = BYTE#47 THEN (* '/' TagTerm *)
// 					mode := 300; (* End Element Section *)
// 				ELSIF C = BYTE#33 THEN (* '!' for Special Section *)
// 					index := index + 1;
// 					mode := 500;
// 				ELSE
// 					s1 := index;
// 				END_IF;
// 				EXIT;
// 			END_IF;
// 			index := index + 1;
// 		END_WHILE;
//
// 		(* analyse element *)
// 		CTRL.TYP := 0; (* TYP löschen *)
// 		IF s1 > 0 THEN
// 			WHILE (index <= stop AND e1 = 0) DO
// 				c := BUF[index];
// 				(* whitespace zeichen = Element with Attributes *)
// 				IF c <= BYTE#32 THEN
// 					(* suche nächstes druckbares zeichen *)
// 					index2 := index;
// 					WHILE (index2 <= stop) AND (BUF[index2] <= BYTE#32) DO
// 						index2 := index2 + 1;
// 					END_WHILE;
// 					IF BUF[index2] = BYTE#47 THEN (* pruefe auf leeres Element '/' *)
// 						index := index2;
// 						e1 := index - 2;
// 						CTRL.TYP := 1; (* struktur-element *)
// 						mode := 300;   (* Close Element *)
// 						EXIT;
// 					END_IF;
//
// 					e1 := index - 1;
// 					CTRL.TYP := 1; (* Element mit Attribute *)
// 					mode := 400;
//
// 				ELSIF c = BYTE#62 THEN (* '>' TagEnd *)
//
// 					(* pruefe auf leeres Element <xx/> *)
// 					index2 := index - 1;
// 					IF BUF[index2] = BYTE#47 THEN (* TagTerm '/' *)
// 						e1 := index2 - 1;
// 						CTRL.TYP := 1;
// 						EMPTY_TAG := TRUE; (* EMPTY TAG Mode *)
// 						mode := 200; (* TEXT Element *)
// 						EXIT;
// 					END_IF;
//
// 					e1 := index - 1;
// 					index2 := index + 1;
//
// 					(* untersuche nachfolgendes Element *)
// 					WHILE (index2 <= stop) DO
// 						c := BUF[index2];
// 						IF c = BYTE#60 THEN (* '<' TagBegin *)
//
// 							index2 := index2 + 1; (* geht bei PCWORX leider nicht anders !*)
// 							c := BUF[index2];
// 							index2 := index2 - 1;
// 							IF c = BYTE#47 THEN (* TagTerm '/' *)
// 								empty_tag := TRUE;
// 								mode := 200; (* TEXT Element *)
// 							ELSE
// 								mode := 100; (* Element *)
// 							END_IF;
// 							CTRL.TYP := 1; (* struktur-element *)
// 							EXIT;
// 						ELSIF c > BYTE#32  THEN (* Printable-Character *)
// 							CTRL.TYP := 1; (* element with text *)
// 							mode := 200;
// 							EXIT;
// 						END_IF;
// 						index2 := index2 + 1;
// 					END_WHILE;
// 				END_IF;
// 				index := index + 1;
// 			END_WHILE;
// 		END_IF;
//
// 		(* Neues Element gefunden*)
// 		IF CTRL.TYP > 0 THEN
//
// 			(* Sonderprüfung auf Processing Instruction (PI) *)
// 			IF BUF[s1] = BYTE#63 THEN (* '?' for Processing Instruction *)
// 				s1 := s1 + 1; (* führendes '?' auslassen *)
// 				CTRL.TYP := 5;
// 			END_IF;
// 			CTRL.BLOCK1_START := INT_TO_UINT(s1);
// 			CTRL.BLOCK1_STOP  := INT_TO_UINT(e1);
// 			CTRL.ELEMENT := BUFFER_TO_STRING(PT:=ADR(BUF),SIZE:=INT_TO_UINT(stop + 1),START:=CTRL.BLOCK1_START,STOP:=CTRL.BLOCK1_STOP);
// 			CTRL.COUNT := CTRL.COUNT + UINT#1;
// 			CTRL.LEVEL := CTRL.LEVEL + UINT#1;
//
// 			IF path_overflow = FALSE THEN
// 				(* Stringlänge überwachen *)
// 				IF LEN(CTRL.PATH) + LEN(CTRL.ELEMENT) + 1 > 250 THEN
// 					path_overflow := TRUE;
// 					CTRL.PATH := 'OVERFLOW';
// 				ELSE
// 					CTRL.PATH := CONCAT(CTRL.PATH,'/');
// 					CTRL.PATH  := CONCAT(CTRL.PATH,CTRL.ELEMENT);
// 				END_IF;
// 			END_IF;
//
// 			IF BIT_OF_DWORD(WORD_TO_DWORD(COMMAND),CTRL.TYP) THEN
//         				(*####################  DEBUG-MESSAGE  ###################################*)
//         				(*IF _debug_enable THEN
//           				LOG_CL.NEW_MSG := 'EL: #T:~1 #C:~2 #E:~3 #P:~6 #L:~7';
//           				LOG_CL.PRINTF[1] := INT_TO_STRING(CTRL.TYP);
//           				LOG_CL.PRINTF[2] := UINT_TO_STRING(CTRL.COUNT);
//           				LOG_CL.PRINTF[3] := CTRL.ELEMENT;
//           				LOG_CL.PRINTF[6] := CTRL.PATH;
//           				LOG_CL.PRINTF[7] := UINT_TO_STRING(CTRL.LEVEL);
//           				LOG_MSG();
//         				END_IF;*)
//         				(*########################################################################*)
// 				RETURN;
// 			END_IF;
// 		END_IF;
//
// 	200: (* ---------- TEXT SECTION ------------------ *)
// 		CTRL.VALUE := '';
// 		IF empty_tag = FALSE THEN
// 			s1 := index;
// 			(* suche '<' EndTag*)
// 			WHILE (index <= stop) AND (BUF[index] <> BYTE#60) DO
// 				index := index + 1;
// 			END_WHILE;
//
// 			E1 := index - 1;
// 			CTRL.BLOCK1_START := INT_TO_UINT(s1);
// 			CTRL.BLOCK1_STOP  := INT_TO_UINT(e1);
// 			CTRL.VALUE := BUFFER_TO_STRING(PT:=ADR(BUF),SIZE:=INT_TO_UINT(stop + 1),START:=CTRL.BLOCK1_START,STOP:=CTRL.BLOCK1_STOP);
// 		END_IF;
//
// 		empty_tag := FALSE;
// 		mode := 300; (* -> NEXT-JOB: END ELEMENT *)
// 		CTRL.COUNT := CTRL.COUNT + UINT#1;
// 		CTRL.TYP := 3;
//
// 		IF BIT_OF_DWORD(WORD_TO_DWORD(command),CTRL.TYP) THEN
//       			(*####################  DEBUG-MESSAGE  ###################################*)
//       			(*IF _debug_enable THEN
//         				LOG_CL.NEW_MSG := 'TE: #T:~1 #C:~2 #E:~3 #V:~4 #P:~6 #L:~7';
//         				LOG_CL.PRINTF[1] := INT_TO_STRING(CTRL.TYP);
//         				LOG_CL.PRINTF[2] := UINT_TO_STRING(CTRL.COUNT);
//         				LOG_CL.PRINTF[3] := CTRL.ELEMENT;
//         				LOG_CL.PRINTF[4] := CTRL.VALUE;
//         				LOG_CL.PRINTF[6] := CTRL.PATH;
//         				LOG_CL.PRINTF[7] := UINT_TO_STRING(CTRL.LEVEL);
//         				LOG_MSG();
//       			END_IF;*)
//       			(*########################################################################*)
// 			RETURN;
// 		END_IF;
//
// 	300: (* ---------- END ELEMENT SECTION ------------------ *)
// 		WHILE (index <= stop) DO
// 			c := BUF[index];
// 			IF c = BYTE#62 THEN (* '>' TagEnd *)
// 				index := index + 1;
// 				s1 := FINDB(str1:=CTRL.PATH,str2:='/');
// 				IF path_overflow = FALSE THEN
// 					IF s1 > 1 THEN
// 						CTRL.ELEMENT := RIGHT(CTRL.PATH,LEN(CTRL.PATH) - s1);
// 						CTRL.PATH := LEFT(CTRL.PATH,s1 - 1);
// 					ELSE
// 						CTRL.ELEMENT := RIGHT(CTRL.PATH,LEN(CTRL.PATH) - 1);
// 						CTRL.PATH :='';
// 					END_IF;
// 				END_IF;
//
// 				CTRL.LEVEL := CTRL.LEVEL - UINT#1;
// 				CTRL.COUNT := CTRL.COUNT + UINT#1;
// 				CTRL.TYP := 2;
// 				mode := 100;
//
// 				IF BIT_OF_DWORD(WORD_TO_DWORD(COMMAND),CTRL.TYP) THEN
//          	 				(*####################  DEBUG-MESSAGE  ###################################*)
//           				(*IF _debug_enable THEN
//             					LOG_CL.NEW_MSG := 'CE: #T:~1 #C:~2 #E:~3 #P:~6 #L:~7';
//             					LOG_CL.PRINTF[1] := INT_TO_STRING(CTRL.TYP);
//             					LOG_CL.PRINTF[2] := UINT_TO_STRING(CTRL.COUNT);
//             					LOG_CL.PRINTF[3] := CTRL.ELEMENT;
//             					LOG_CL.PRINTF[6] := CTRL.PATH;
//             					LOG_CL.PRINTF[7] := UINT_TO_STRING(CTRL.LEVEL);
//             					LOG_MSG();
//           				END_IF;*)
//           				(*########################################################################*)
// 					RETURN;
// 				ELSE
// 					EXIT;
// 				END_IF;
// 			END_IF;
// 			index := index + 1;
// 		END_WHILE;
//
// 	400: (* ---------- ATTRIBUTE SECTION ------------------ *)
// 		(* search first normal charakter *)
// 		WHILE (index <= stop AND BUF[index] <= BYTE#32) DO
// 			index := index + 1;
// 		END_WHILE;
//
// 		(* begin Attribe name *)
// 		e1 := 0;
// 		s1 := index;
// 		(* search end of Attrib Name '=' *)
// 		WHILE (index <= stop) DO
// 			IF BUF[index] = BYTE#61 THEN (* '=' Equals *)
// 				e1 := index - 1;
// 				EXIT;
// 			END_IF;
// 			index := index + 1;
// 		END_WHILE;
//
// 		IF e1 > 0 THEN
// 			(* Attribute Name *)
// 			CTRL.BLOCK1_START := INT_TO_UINT(s1);
// 			CTRL.BLOCK1_STOP  := INT_TO_UINT(e1);
// 			CTRL.ATTRIBUTE := BUFFER_TO_STRING(PT:=ADR(BUF),SIZE:=INT_TO_UINT(STOP + 1),START:=CTRL.BLOCK1_START,STOP:=CTRL.BLOCK1_STOP);
// 			(* search end of Attrib Value '=' *)
// 			index := index + 2;
// 			e1 := 0;
// 			s1 := INDEX;
// 			WHILE (index <= stop AND e1 = 0) DO
// 				c := BUF[index];
// 				IF c = BYTE#34 OR c = BYTE#39 THEN (* " OR ' Equals *)
// 					e1 := index - 1;
// 				END_IF;
// 				index := index + 1;
// 			END_WHILE;
//
// 			IF e1 > 0 THEN
// 				(* Value *)
// 				CTRL.BLOCK2_START := INT_TO_UINT(s1);
// 				CTRL.BLOCK2_STOP  := INT_TO_UINT(e1);
//
// 				(* bei leeren "" ist start groesser als stop und wird somit zum leerstring *)
// 				CTRL.VALUE := BUFFER_TO_STRING(PT:=ADR(BUF),SIZE:=INT_TO_UINT(stop + 1),START:=CTRL.BLOCK2_START,STOP:=CTRL.BLOCK2_STOP);
// 				(* search next non white space charakter *)
// 				WHILE (index <= stop AND BUF[index] <= BYTE#32) DO
// 					index := index + 1;
// 				END_WHILE;
//
// 					c := BUF[index];
// 					(* TagEnd '>' *)
// 					IF c = BYTE#62 THEN
// 						index := index + 1;
// 						index2 := index;
//
// 					(* search next non white space charakter *)
// 					WHILE (index <= stop AND BUF[index] <= BYTE#32) DO
// 						index := index + 1;
// 					END_WHILE;
//
// 					IF BUF[index] = BYTE#60 THEN (* TagBegin '<' *)
// 						mode := 100; (* -> NEXT-JOB: ELEMENT-SECTION *)
// 					ELSE
// 						index := index2;
// 						mode := 200; (* -> NEXT-JOB: TEXT-SECTION *)
// 					END_IF;
//
// 				ELSIF c = BYTE#47 OR c = BYTE#63 THEN (* TagTerm '/' OR '?' end Processing Instruction *)
// 					mode := 300; (* -> NEXT-JOB: END ELEMENT *)
// 				ELSE
// 					mode := 400; (* -> NEXT-JOB: ATTRIBUTE-SECTION *)
// 				END_IF;
//
// 				CTRL.COUNT := CTRL.COUNT + UINT#1;
// 				CTRL.TYP := 4;
// 				IF BIT_OF_DWORD(WORD_TO_DWORD(command),CTRL.TYP) THEN
//           				(*####################  DEBUG-MESSAGE  ###################################*)
//           				(*IF _debug_enable THEN
//             					LOG_CL.NEW_MSG := 'AT: #T:~1 #C:~2 #E:~3 #A:~4 #V:~5 #P:~6 #L:~7';
//             					LOG_CL.PRINTF[1] := INT_TO_STRING(CTRL.TYP);
//             					LOG_CL.PRINTF[2] := UINT_TO_STRING(CTRL.COUNT);
//             					LOG_CL.PRINTF[3] := CTRL.ELEMENT;
//             					LOG_CL.PRINTF[4] := CTRL.ATTRIBUTE;
//             					LOG_CL.PRINTF[5] := CTRL.VALUE;
//             					LOG_CL.PRINTF[6] := CTRL.PATH;
//             					LOG_CL.PRINTF[7] := UINT_TO_STRING(CTRL.LEVEL);
//             					LOG_MSG();
//           				END_IF;*)
//           				(*########################################################################*)
// 					RETURN;
// 				END_IF;
// 			END_IF;
// 		END_IF;
//
// 	500: (* ---------- SPECIAL DATA SECTION (Document Type Declarations) ---------- *)
//
// 		CTRL.TYP := 0;
// 		s1 := 0;
// 		index2 := 11;
//
// 		WHILE (s1 = 0) DO
// 			index2 := index2 + 1;
// 			CTRL.TYP := index2;
//
// 			CASE index2 OF
// 			12: (* CDATA *)
// 				s_code := '[CDATA[';
// 				e_code := ']]>';
// 			13: (* COMMENT *)
// 				s_code := '--';
// 				e_code := '-->';
// 			14: (* ANY DTD *)
// 				e_code := '';
// 				s1 := index;
// 				EXIT;
// 			END_CASE;
//
// 			e1 := LEN(s_code);
// 			IF BUFFER_SEARCH(PT:=ADR(BUF),SIZE:=INT_TO_UINT(index + e1),STR:=S_CODE,POS:=index,IGN:=FALSE) = INDEX THEN
// 				s1 := index + e1;
// 			END_IF;
// 		END_WHILE;
//
// 		CTRL.BLOCK1_START := INT_TO_UINT(s1);
// 		IF LEN(e_code) > 0 THEN
// 			(* Ende Kennung suchen *)
// 			e1 := BUFFER_SEARCH(PT:=ADR(BUF),SIZE:=INT_TO_UINT(stop + 1),STR:=e_code,POS:=index,IGN:=FALSE);
// 			CTRL.BLOCK1_STOP := INT_TO_UINT(e1 - 1);
// 			index := e1 + LEN(e_code); (* naechstes element *)
// 		ELSE
// 			(* suche '>' EndTag*)
// 			index2 := 1; (* <> Paar zähler *)
// 			WHILE (index <= stop AND index2 > 0) DO
// 				c := BUF[index];
// 				IF c = BYTE#60 THEN (* '<' TagBegin *)
// 					index2 := index2 + 1;
// 				ELSIF c = BYTE#62 THEN (* '>' TagEnd   *)
// 					index2 := index2 - 1;
// 				ELSIF c = BYTE#34 OR c = BYTE#39 THEN (* " Double Quote OR ' Single Quote *)
// 					index := index + 1;
// 					WHILE (index <= stop) DO
// 						c := BUF[index];
// 						IF c = BYTE#34 OR c = BYTE#39 THEN (* " Double Quote OR ' Single Quote *)
// 							EXIT;
// 						END_IF;
// 						index := index + 1;
// 					END_WHILE;
// 				END_IF;
// 				index := index + 1;
// 			END_WHILE;
// 			CTRL.BLOCK1_STOP := INT_TO_UINT(index - 2);
// 		END_IF;
//
// 		CTRL.VALUE := BUFFER_TO_STRING(PT:=ADR(BUF),SIZE:=INT_TO_UINT(stop + 1),START:=CTRL.BLOCK1_START,STOP:=CTRL.BLOCK1_STOP);
// 		CTRL.COUNT := CTRL.COUNT + UINT#1;
// 		mode := 100; (* -> NEXT-JOB: ELEMENT *)
//
// 		IF BIT_OF_DWORD(WORD_TO_DWORD(command),CTRL.TYP) THEN
//       			(*####################  DEBUG-MESSAGE  ###################################*)
//       			(*IF _debug_enable THEN
//         				LOG_CL.NEW_MSG := 'DTD: #T:~1 #C:~2 #S:~3 #E:~4 #V:~5 #P:~6 #L:~7';
//         				LOG_CL.PRINTF[1] := INT_TO_STRING(CTRL.TYP);
//         				LOG_CL.PRINTF[2] := UINT_TO_STRING(CTRL.COUNT);
//         				LOG_CL.PRINTF[3] := UINT_TO_STRING(CTRL.BLOCK1_START);
//         				LOG_CL.PRINTF[4] := UINT_TO_STRING(CTRL.BLOCK1_STOP);
//         				LOG_CL.PRINTF[5] := CTRL.VALUE;
//         				LOG_CL.PRINTF[6] := CTRL.PATH;
//         				LOG_CL.PRINTF[7] := UINT_TO_STRING(CTRL.LEVEL);
//         				LOG_MSG();
//       			END_IF;*)
//       			(*########################################################################*)
// 			RETURN;
// 		END_IF;
//
// 	END_CASE;
// END_WHILE;
// END_FUNCTION_BLOCK
